(* Logix 5000 project; controller TFF vendor 1 type 14 code 107 rev 33.11; software revision 33.04; part 21 of 38 *)
(* tags used below, declared in another part *)
   Config : Configuration;   // Index Array used in configuration routines
   TIME : DINT[2];
   AA008 : ALIAS FOR DigitalPoint[18];
   AI101_SIG : ALIAS FOR DigitalPoint[106];
   AI104_SIG : ALIAS FOR DigitalPoint[107];
   AI201A_SIG : ALIAS FOR DigitalPoint[90];
   AI201B_SIG : ALIAS FOR DigitalPoint[109];
   AI202_SIG : ALIAS FOR DigitalPoint[105];
   AI203_SIG : ALIAS FOR DigitalPoint[91];
   AI204_SIG : ALIAS FOR DigitalPoint[92];
   DF24VDC : ALIAS FOR DigitalPoint[4];
   DF24VDCPC : ALIAS FOR DigitalPoint[25];
   DF3PHP003 : ALIAS FOR DigitalPoint[27];
   DF48MIX : ALIAS FOR DigitalPoint[26];
   DF48P001 : ALIAS FOR DigitalPoint[23];
   DF48P002 : ALIAS FOR DigitalPoint[24];
   Diafiltration : Diafiltration;
   DigitalPoint : DigitalPoint[150];   // Digital Point Array
   Drive : Drive[11];   // Drives Array
   ES001 : ALIAS FOR DigitalPoint[2];
   ExternalTCU : BOOL;   // Use of External TCU
   ExternalWeight : BOOL;   // Use of External Weight
   FI101_SIG : ALIAS FOR DigitalPoint[110];
   FI201_SIG : ALIAS FOR DigitalPoint[93];
   FI401_SIG : ALIAS FOR DigitalPoint[94];
   FlowPath : FlowPath[64];   // Flow Path Array
   FlowPathControl : FlowPathControl;   // Flow Path Control
   Gateway : Gateway;   // Gateway Control
   MIX101 : ALIAS FOR AnalogPoint[14];
   MIX101_SIG : ALIAS FOR DigitalPoint[104];
   MIX101DF : ALIAS FOR DigitalPoint[28];
   Mixer : Mixer;   // Mixer config. structure
   Options : Options;   // Options List
   PCV101 : ALIAS FOR AnalogPoint[3];
   PCV101_SIG : ALIAS FOR DigitalPoint[102];
   PCV201 : ALIAS FOR AnalogPoint[4];
   PCV201_SIG : ALIAS FOR DigitalPoint[103];
   PI001_SIG : ALIAS FOR DigitalPoint[97];
   PI101_SIG : ALIAS FOR DigitalPoint[98];
   PI201_SIG : ALIAS FOR DigitalPoint[99];
   PI401_SIG : ALIAS FOR DigitalPoint[100];
   PI601_SIG : ALIAS FOR DigitalPoint[95];
   PISL601 : ALIAS FOR DigitalPoint[0];
   PISL602 : ALIAS FOR DigitalPoint[1];
   PSH001 : ALIAS FOR DigitalPoint[21];
   PSH401 : ALIAS FOR DigitalPoint[22];
   RSBUZZ : ALIAS FOR DigitalPoint[3];
   SIC001 : ALIAS FOR Drive[1];
   SIC001DF : ALIAS FOR DigitalPoint[16];
   SIC002 : ALIAS FOR Drive[2];
   SIC002DF : ALIAS FOR DigitalPoint[17];
   SIC003DF : ALIAS FOR DigitalPoint[29];
   SIC004 : ALIAS FOR Drive[3];
   Tank : TankManagement;   // Tank Management
   TCU101_SIG : ALIAS FOR DigitalPoint[108];
   TCU101DF : ALIAS FOR DigitalPoint[30];
   TI101_SIG : ALIAS FOR DigitalPoint[101];
   TI201_SIG : ALIAS FOR DigitalPoint[111];
   UserCr1 : ALIAS FOR DigitalPoint[65];
   UserCr2 : ALIAS FOR DigitalPoint[67];
   UserNCr1 : ALIAS FOR DigitalPoint[64];
   UserNCr2 : ALIAS FOR DigitalPoint[66];
   Valve : Valve[100];   // Valve Array
   WI201_SIG : ALIAS FOR DigitalPoint[96];
   XS011 : ALIAS FOR DigitalPoint[14];
   XS012 : ALIAS FOR DigitalPoint[15];
   XV003 : ALIAS FOR Valve[2];
   YA01 : ALIAS FOR DigitalPoint[50];
   YA02 : ALIAS FOR DigitalPoint[51];
   YA03 : ALIAS FOR DigitalPoint[52];
   YA04 : ALIAS FOR DigitalPoint[53];
   YA05 : ALIAS FOR DigitalPoint[54];
   YA06 : ALIAS FOR DigitalPoint[55];
   YA07 : ALIAS FOR DigitalPoint[56];
   YA08 : ALIAS FOR DigitalPoint[57];
   YA09 : ALIAS FOR DigitalPoint[58];
   YA10 : ALIAS FOR DigitalPoint[59];
   YA11 : ALIAS FOR DigitalPoint[60];
   YA12 : ALIAS FOR DigitalPoint[61];
   YA13 : ALIAS FOR DigitalPoint[62];
   YA14 : ALIAS FOR DigitalPoint[63];
   YA15 : ALIAS FOR DigitalPoint[69];
   YA16 : ALIAS FOR DigitalPoint[70];
   YA17 : ALIAS FOR DigitalPoint[71];
   YA18 : ALIAS FOR DigitalPoint[72];
   YA41 : ALIAS FOR DigitalPoint[73];
   ZS001 : ALIAS FOR DigitalPoint[6];
   ZS002 : ALIAS FOR DigitalPoint[7];
   ZS003 : ALIAS FOR DigitalPoint[8];
   ZS004 : ALIAS FOR DigitalPoint[9];
   ZS005 : ALIAS FOR DigitalPoint[10];
   ZS008 : ALIAS FOR DigitalPoint[5];
   ZSDF : ALIAS FOR DigitalPoint[68];
(* Process, continued *)

ROUTINE Config_DigitalPoint_Real   (* structured text *)
// Apply the default configuration
   (* ==========================================================
   	Config DigitalPoint Real : Configure DigitalPoint Structure (for real input)
   
   	List of treatments
   		- DigitalPoint[0] : Valves Air Defect PISL601
   		- DigitalPoint[1] : Manifold Valves Air Defect PISL602
   		- DigitalPoint[2] : Emergency Stop ES001
   		- DigitalPoint[3] : Reset Buzzer RSBUZZ
   		- DigitalPoint[4] : 24 VDC defect DF24VDC
   		- DigitalPoint[5] : Door Closed ZS008
   		- DigitalPoint[6] : Clamshell Locking 1 Closed ZS001
   		- DigitalPoint[7] : Clamshell Locking 2 Closed ZS002
   		- DigitalPoint[8] : Clamshell Locking 3 Closed ZS003
   		- DigitalPoint[9] : Clamshell Locking 4 Closed ZS004
   		- DigitalPoint[10]: Clamshell Locking 5 Closed ZS005
   		- Reset Loop : Set to 0 the DigitalPoint[11 to 13].EnableCfg
   		- DigitalPoint[14]: Pump P001 Type XS011
   		- DigitalPoint[15]: Pump P002 Type XS012
   		- DigitalPoint[16]: P001 Defect SIC001DF
   		- DigitalPoint[17]: P002 Defect SIC002DF
   		- DigitalPoint[18]: C8000 Defect AA008
   		- DigitalPoint[19]: Spare
   		- DigitalPoint[20]: Spare
   		- DigitalPoint[21]: Feed Pump High Pressure PSH001
   		- DigitalPoint[22]: Transfer Pump High Pressure PSH401
   		- DigitalPoint[23]: P001 48 VDC Defect DF48P001
   		- DigitalPoint[24]: P002 48 VDC Defect DF48P002
   		- DigitalPoint[25]: Pump Cart 24 VDC Defect DF24VDCPC
   		- DigitalPoint[26]: Mixer 48 VDC Defect DF48MIX
   		- DigitalPoint[27]: Pump P003 Power Supply Defect DF3PHP003
   		- DigitalPoint[28]: Mixer Defect MIX101DF
   		- DigitalPoint[29]: P003 Defect SIC003DF
   		- DigitalPoint[30]: TCU Defect TCU101DF
   		- Reset Loop : Set to 0 the DigitalPoint[31 to 33].EnableCfg
   		- DigitalPoint[34]: Exchange DI#1
   		- DigitalPoint[35]: Exchange DI#2
   		- DigitalPoint[36]: Exchange DI#3
   		- DigitalPoint[37]: Exchange DI#4
   		- DigitalPoint[38]: Exchange DI#5
   		- DigitalPoint[39]: Exchange DI#6
   		- DigitalPoint[40]: Exchange DI#7
   		- DigitalPoint[41]: Exchange DI#8
   		- Reset Loop : Set to 0 the DigitalPoint[42 to 49].EnableCfg
   
   -----------------------------------------------------------------------------------------------------------------------------------------------------
   	History
   		2019-DEC-24 - Merck - Q. Spindler - Initial version for Candidate Release 1.00.00.00.a
   		2020-MAR-27 - Merck - Q. Spindler - Modifications for Candidate Release 1.00.00.00.b
   					- Add Options for AA008
   		2020-SEP-09 - Merck - Q. Spindler - Modifications for Candidate Release 1.00.00.00.d
   					- Change PriorityCfg to 0 and set Priority to 1 for PSH001 and PSH401
   					- Disable TCU101DF alarm if ExternalTCU not used
   ============================================================*)
   
   (*DigitalPoint[0] : Valves Air Defect PISL601
   ============================================================*)
   DigitalPoint[0].EnableCfg := 1 ;
   DigitalPoint[0].ActiveStateCFg := 1 ;
   DigitalPoint[0].RealInputCfg := 1 ;
   DigitalPoint[0].InputAddressCfg := 0 ;
   DigitalPoint[0].AlarmCfg := 1 ;
   DigitalPoint[0].AlarmStateCfg := 0 ;
   DigitalPoint[0].OverrideCfg := 1 ;
   DigitalPoint[0].PriorityCfg := 1 ;
   DigitalPoint[0].Cond1Cfg := 0 ;
   DigitalPoint[0].Cond2Cfg := 0 ;
   DigitalPoint[0].FlashingInputCfg := 0 ;
   
   (*DigitalPoint[1] : Manifold Valves Air Defect PISL602
   ============================================================*)
   DigitalPoint[1].EnableCfg := 1 ;
   DigitalPoint[1].ActiveStateCFg := 1 ;
   DigitalPoint[1].RealInputCfg := 1 ;
   DigitalPoint[1].InputAddressCfg := 1 ;
   DigitalPoint[1].AlarmCfg := 1 ;
   DigitalPoint[1].AlarmStateCfg := 0 ;
   DigitalPoint[1].OverrideCfg := 1 ;
   DigitalPoint[1].PriorityCfg := 1 ;
   DigitalPoint[1].Cond1Cfg := 0 ;
   DigitalPoint[1].Cond2Cfg := 0 ;
   DigitalPoint[1].FlashingInputCfg := 0 ;
   
   (*DigitalPoint[2] : Emergency Stop ES001
   ============================================================*)
   DigitalPoint[2].EnableCfg := 1 ;
   DigitalPoint[2].ActiveStateCFg := 1 ;
   DigitalPoint[2].RealInputCfg := 1 ;
   DigitalPoint[2].InputAddressCfg := 2 ;
   DigitalPoint[2].AlarmCfg := 1 ;
   DigitalPoint[2].AlarmStateCfg := 0 ;
   DigitalPoint[2].OverrideCfg := 0 ;
   DigitalPoint[2].PriorityCfg := 0 ;
   DigitalPoint[2].Priority := 1 ;
   DigitalPoint[2].Cond1Cfg := 0 ;
   DigitalPoint[2].Cond2Cfg := 0 ;
   DigitalPoint[2].FlashingInputCfg := 0 ;
   
   (*DigitalPoint[3] : Reset Buzzer RSBUZZ
   ============================================================*)
   DigitalPoint[3].EnableCfg := 1 ;
   DigitalPoint[3].ActiveStateCFg := 1 ;
   DigitalPoint[3].RealInputCfg := 1 ;
   DigitalPoint[3].InputAddressCfg := 3 ;
   DigitalPoint[3].AlarmCfg := 0 ;
   DigitalPoint[3].Alarm := 0 ;
   DigitalPoint[3].AlarmStateCfg := 0 ;
   DigitalPoint[3].OverrideCfg := 0 ;
   DigitalPoint[3].Priority := 0 ;
   DigitalPoint[3].PriorityCfg := 0 ;
   DigitalPoint[3].Cond1Cfg := 0 ;
   DigitalPoint[3].Cond2Cfg := 0 ;
   DigitalPoint[3].FlashingInputCfg := 0 ;
   
   (*DigitalPoint[4] : 24 VDC defect DF24VDC
   ============================================================*)
   DigitalPoint[4].EnableCfg := 1 ;
   DigitalPoint[4].ActiveStateCFg := 1 ;
   DigitalPoint[4].RealInputCfg := 1 ;
   DigitalPoint[4].InputAddressCfg := 4 ;
   DigitalPoint[4].AlarmCfg := 1 ;
   DigitalPoint[4].AlarmStateCfg := 0 ;
   DigitalPoint[4].OverrideCfg := 1 ;
   DigitalPoint[4].PriorityCfg := 1 ;
   DigitalPoint[4].Cond1Cfg := 0 ;
   DigitalPoint[4].Cond2Cfg := 0 ;
   DigitalPoint[4].FlashingInputCfg := 0 ;
   
   (*DigitalPoint[5] : Door Closed ZS008
   ============================================================*)
   DigitalPoint[5].EnableCfg := 1 ;
   DigitalPoint[5].ActiveStateCFg := 1 ;
   DigitalPoint[5].RealInputCfg := 1 ;
   DigitalPoint[5].InputAddressCfg := 5 ;
   DigitalPoint[5].AlarmCfg := 1 ;
   DigitalPoint[5].AlarmStateCfg := 0 ;
   DigitalPoint[5].OverrideCfg := 1 ;
   DigitalPoint[5].PriorityCfg := 1 ;
   DigitalPoint[5].Cond1Cfg := 0 ;
   DigitalPoint[5].Cond2Cfg := 0 ;
   DigitalPoint[5].FlashingInputCfg := 0 ;
   
   (*DigitalPoint[6] : Clamshell Locking 1 Closed ZS001
   ============================================================*)
   DigitalPoint[6].EnableCfg := 1 ;
   DigitalPoint[6].ActiveStateCFg := 1 ;
   DigitalPoint[6].RealInputCfg := 1 ;
   DigitalPoint[6].InputAddressCfg := 6 ;
   DigitalPoint[6].AlarmCfg := 0 ;
   DigitalPoint[6].Alarm := 0 ;
   DigitalPoint[6].AlarmStateCfg := 0 ;
   DigitalPoint[6].OverrideCfg := 0 ;
   DigitalPoint[6].PriorityCfg := 0 ;
   DigitalPoint[6].Cond1Cfg := 0 ;
   DigitalPoint[6].Cond2Cfg := 0 ;
   DigitalPoint[6].FlashingInputCfg := 0 ;
   
   (*DigitalPoint[7] : Clamshell Locking 2 Closed ZS002
   ============================================================*)
   DigitalPoint[7].EnableCfg := 1 ;
   DigitalPoint[7].ActiveStateCFg := 1 ;
   DigitalPoint[7].RealInputCfg := 1 ;
   DigitalPoint[7].InputAddressCfg := 7 ;
   DigitalPoint[7].AlarmCfg := 0 ;
   DigitalPoint[7].Alarm := 0 ;
   DigitalPoint[7].AlarmStateCfg := 0 ;
   DigitalPoint[7].OverrideCfg := 0 ;
   DigitalPoint[7].PriorityCfg := 0 ;
   DigitalPoint[7].Cond1Cfg := 0 ;
   DigitalPoint[7].Cond2Cfg := 0 ;
   DigitalPoint[7].FlashingInputCfg := 0 ;
   
   (*DigitalPoint[8] : Clamshell Locking 3 Closed ZS003
   ============================================================*)
   DigitalPoint[8].EnableCfg := 1 ;
   DigitalPoint[8].ActiveStateCFg := 1 ;
   DigitalPoint[8].RealInputCfg := 1 ;
   DigitalPoint[8].InputAddressCfg := 8 ;
   DigitalPoint[8].AlarmCfg := 0 ;
   DigitalPoint[8].Alarm := 0 ;
   DigitalPoint[8].AlarmStateCfg := 0 ;
   DigitalPoint[8].OverrideCfg := 0 ;
   DigitalPoint[8].PriorityCfg := 0 ;
   DigitalPoint[8].Cond1Cfg := 0 ;
   DigitalPoint[8].Cond2Cfg := 0 ;
   DigitalPoint[8].FlashingInputCfg := 0 ;
   
   (*DigitalPoint[9] : Clamshell Locking 4 Closed ZS004
   ============================================================*)
   DigitalPoint[9].EnableCfg := 1 ;
   DigitalPoint[9].ActiveStateCFg := 1 ;
   DigitalPoint[9].RealInputCfg := 1 ;
   DigitalPoint[9].InputAddressCfg := 9 ;
   DigitalPoint[9].AlarmCfg := 0 ;
   DigitalPoint[9].Alarm := 0 ;
   DigitalPoint[9].AlarmStateCfg := 0 ;
   DigitalPoint[9].OverrideCfg := 0 ;
   DigitalPoint[9].PriorityCfg := 0 ;
   DigitalPoint[9].Cond1Cfg := 0 ;
   DigitalPoint[9].Cond2Cfg := 0 ;
   DigitalPoint[9].FlashingInputCfg := 0 ;
   
   (*DigitalPoint[10]: Clamshell Locking 5 Closed ZS005
   ============================================================*)
   DigitalPoint[10].EnableCfg := 1 ;
   DigitalPoint[10].ActiveStateCFg := 1 ;
   DigitalPoint[10].RealInputCfg := 1 ;
   DigitalPoint[10].InputAddressCfg := 10 ;
   DigitalPoint[10].AlarmCfg := 0 ;
   DigitalPoint[10].Alarm := 0 ;
   DigitalPoint[10].AlarmStateCfg := 0 ;
   DigitalPoint[10].OverrideCfg := 0 ;
   DigitalPoint[10].PriorityCfg := 0 ;
   DigitalPoint[10].Cond1Cfg := 0 ;
   DigitalPoint[10].Cond2Cfg := 0 ;
   DigitalPoint[10].FlashingInputCfg := 0 ;
   
   
   (*Reset Loop : Set to 0 the DigitalPoint[11 to 13].EnableCfg
   ============================================================*)
   FOR Config.IndexDP := 11 to 13 do
   	DigitalPoint[Config.IndexDP].EnableCfg := 0 ;
   	DigitalPoint[Config.IndexDP].AlarmCfg := 0 ;
   	DigitalPoint[Config.IndexDP].Alarm := 0 ;
   End_for ;
   
   
   (*DigitalPoint[14]: Pump P001 Type XS011
   ============================================================*)
   DigitalPoint[14].EnableCfg := 1 ;
   DigitalPoint[14].ActiveStateCFg := 1 ;
   DigitalPoint[14].RealInputCfg := 1 ;
   DigitalPoint[14].InputAddressCfg := 14 ;
   DigitalPoint[14].AlarmCfg := 0 ;
   DigitalPoint[14].Alarm := 0 ;
   DigitalPoint[14].AlarmStateCfg := 0 ;
   DigitalPoint[14].OverrideCfg := 0 ;
   DigitalPoint[14].PriorityCfg := 0 ;
   DigitalPoint[14].Cond1Cfg := 0 ;
   DigitalPoint[14].Cond2Cfg := 0 ;
   DigitalPoint[14].FlashingInputCfg := 0 ;
   
   (*DigitalPoint[15]: Pump P002 Type XS012
   ============================================================*)
   DigitalPoint[15].EnableCfg := 1 ;
   DigitalPoint[15].ActiveStateCFg := 1 ;
   DigitalPoint[15].RealInputCfg := 1 ;
   DigitalPoint[15].InputAddressCfg := 15 ;
   DigitalPoint[15].AlarmCfg := 0 ;
   DigitalPoint[15].Alarm := 0 ;
   DigitalPoint[15].AlarmStateCfg := 0 ;
   DigitalPoint[15].OverrideCfg := 0 ;
   DigitalPoint[15].PriorityCfg := 0 ;
   DigitalPoint[15].Cond1Cfg := 0 ;
   DigitalPoint[15].Cond2Cfg := 0 ;
   DigitalPoint[15].FlashingInputCfg := 0 ;
   
   (*DigitalPoint[16]: P001 Defect SIC001DF
   ============================================================*)
   DigitalPoint[16].EnableCfg := 1 ;
   DigitalPoint[16].ActiveStateCFg := 1 ;
   DigitalPoint[16].RealInputCfg := 1 ;
   DigitalPoint[16].InputAddressCfg := 16 ;
   DigitalPoint[16].AlarmCfg := 1 ;
   DigitalPoint[16].AlarmStateCfg := 0 ;
   DigitalPoint[16].OverrideCfg := 1 ;
   DigitalPoint[16].PriorityCfg := 1 ;
   DigitalPoint[16].Cond1Cfg := 0 ;
   DigitalPoint[16].Cond2Cfg := 0 ;
   DigitalPoint[16].FlashingInputCfg := 0 ;
   
   (*DigitalPoint[17]: P002 Defect SIC002DF
   ============================================================*)
   DigitalPoint[17].EnableCfg := 1 ;
   DigitalPoint[17].ActiveStateCFg := 1 ;
   DigitalPoint[17].RealInputCfg := 1 ;
   DigitalPoint[17].InputAddressCfg := 17 ;
   DigitalPoint[17].AlarmCfg := 1 ;
   DigitalPoint[17].AlarmStateCfg := 0 ;
   DigitalPoint[17].OverrideCfg := 1 ;
   DigitalPoint[17].PriorityCfg := 1 ;
   DigitalPoint[17].Cond1Cfg := 0 ;
   DigitalPoint[17].Cond2Cfg := 0 ;
   DigitalPoint[17].FlashingInputCfg := 0 ;
   
   (*DigitalPoint[18]: C8000 Defect AA008
   ============================================================*)
   If Options.FiltrateCondPHUV OR Options.FiltrateCondPH Then
   	DigitalPoint[18].EnableCfg := 1 ;
   	DigitalPoint[18].AlarmCfg := 1 ;
   Else
   	DigitalPoint[18].EnableCfg := 0 ;
   	DigitalPoint[18].AlarmCfg := 0 ;
   	DigitalPoint[18].Alarm := 0 ;
   End_if;
   
   DigitalPoint[18].ActiveStateCFg := 1 ;
   DigitalPoint[18].RealInputCfg := 1 ;
   DigitalPoint[18].InputAddressCfg := 18 ;
   DigitalPoint[18].AlarmStateCfg := 0 ;
   DigitalPoint[18].OverrideCfg := 1 ;
   DigitalPoint[18].PriorityCfg := 1 ;
   DigitalPoint[18].Cond1Cfg := 0 ;
   DigitalPoint[18].Cond2Cfg := 0 ;
   DigitalPoint[18].FlashingInputCfg := 0 ;
   
   (*DigitalPoint[19]: Spare
   ============================================================*)
   DigitalPoint[19].EnableCfg := 0 ;
   DigitalPoint[19].ActiveStateCFg := 1 ;
   DigitalPoint[19].RealInputCfg := 1 ;
   DigitalPoint[19].InputAddressCfg := 19 ;
   DigitalPoint[19].AlarmCfg := 0 ;
   DigitalPoint[19].AlarmStateCfg := 0 ;
   DigitalPoint[19].OverrideCfg := 1 ;
   DigitalPoint[19].PriorityCfg := 1 ;
   DigitalPoint[19].Cond1Cfg := 0 ;
   DigitalPoint[19].Cond2Cfg := 0 ;
   DigitalPoint[19].FlashingInputCfg := 0 ;
   
   (*DigitalPoint[20]: Spare
   ============================================================*)
   DigitalPoint[20].EnableCfg := 0 ;
   DigitalPoint[20].ActiveStateCFg := 1 ;
   DigitalPoint[20].RealInputCfg := 1 ;
   DigitalPoint[20].InputAddressCfg := 20 ;
   DigitalPoint[20].AlarmCfg := 0 ;
   DigitalPoint[20].AlarmStateCfg := 0 ;
   DigitalPoint[20].OverrideCfg := 1 ;
   DigitalPoint[20].PriorityCfg := 1 ;
   DigitalPoint[20].Cond1Cfg := 0 ;
   DigitalPoint[20].Cond2Cfg := 0 ;
   DigitalPoint[20].FlashingInputCfg := 0 ;
   
   (*DigitalPoint[21]: Feed Pump High Pressure PSH001
   ============================================================*)
   DigitalPoint[21].EnableCfg := 1 ;
   DigitalPoint[21].ActiveStateCFg := 1 ;
   DigitalPoint[21].RealInputCfg := 1 ;
   DigitalPoint[21].InputAddressCfg := 21 ;
   DigitalPoint[21].AlarmCfg := 1 ;
   DigitalPoint[21].AlarmStateCfg := 0 ;
   DigitalPoint[21].OverrideCfg := 1 ;
   DigitalPoint[21].PriorityCfg := 0 ;
   DigitalPoint[21].Priority := 1 ;
   DigitalPoint[21].Cond1Cfg := 0 ;
   DigitalPoint[21].Cond2Cfg := 0 ;
   DigitalPoint[21].FlashingInputCfg := 0 ;
   
   (*DigitalPoint[22]: Transfer Pump High Pressure PSH401
   ============================================================*)
   DigitalPoint[22].EnableCfg := 1 ;
   DigitalPoint[22].ActiveStateCFg := 1 ;
   DigitalPoint[22].RealInputCfg := 1 ;
   DigitalPoint[22].InputAddressCfg := 22 ;
   DigitalPoint[22].AlarmCfg := 1 ;
   DigitalPoint[22].AlarmStateCfg := 0 ;
   DigitalPoint[22].OverrideCfg := 1 ;
   DigitalPoint[22].PriorityCfg := 0 ;
   DigitalPoint[22].Priority := 1 ;
   DigitalPoint[22].Cond1Cfg := 0 ;
   DigitalPoint[22].Cond2Cfg := 0 ;
   DigitalPoint[22].FlashingInputCfg := 0 ;
   
   (*DigitalPoint[23]: P001 48 VDC Defect DF48P001
   ============================================================*)
   DigitalPoint[23].EnableCfg := 1 ;
   DigitalPoint[23].ActiveStateCFg := 1 ;
   DigitalPoint[23].RealInputCfg := 1 ;
   DigitalPoint[23].InputAddressCfg := 23 ;
   DigitalPoint[23].AlarmCfg := 1 ;
   DigitalPoint[23].AlarmStateCfg := 0 ;
   DigitalPoint[23].OverrideCfg := 1 ;
   DigitalPoint[23].PriorityCfg := 1 ;
   DigitalPoint[23].Cond1Cfg := 0 ;
   DigitalPoint[23].Cond2Cfg := 0 ;
   DigitalPoint[23].FlashingInputCfg := 0 ;
   
   (*DigitalPoint[24]: P002 48 VDC Defect DF48P002
   ============================================================*)
   DigitalPoint[24].EnableCfg := 1 ;
   DigitalPoint[24].ActiveStateCFg := 1 ;
   DigitalPoint[24].RealInputCfg := 1 ;
   DigitalPoint[24].InputAddressCfg := 24 ;
   DigitalPoint[24].AlarmCfg := 1 ;
   DigitalPoint[24].AlarmStateCfg := 0 ;
   DigitalPoint[24].OverrideCfg := 1 ;
   DigitalPoint[24].PriorityCfg := 1 ;
   DigitalPoint[24].Cond1Cfg := 0 ;
   DigitalPoint[24].Cond2Cfg := 0 ;
   DigitalPoint[24].FlashingInputCfg := 0 ;
   
   (*DigitalPoint[25]: Pump Cart 24 VDC Defect DF24VDCPC
   ============================================================*)
   DigitalPoint[25].EnableCfg := 1 ;
   DigitalPoint[25].ActiveStateCFg := 1 ;
   DigitalPoint[25].RealInputCfg := 1 ;
   DigitalPoint[25].InputAddressCfg := 25 ;
   DigitalPoint[25].AlarmCfg := 1 ;
   DigitalPoint[25].AlarmStateCfg := 0 ;
   DigitalPoint[25].OverrideCfg := 1 ;
   DigitalPoint[25].PriorityCfg := 1 ;
   DigitalPoint[25].Cond1Cfg := 0 ;
   DigitalPoint[25].Cond2Cfg := 0 ;
   DigitalPoint[25].FlashingInputCfg := 0 ;
   
   (*DigitalPoint[26]: Mixer 48 VDC Defect DF48MIX
   ============================================================*)
   (*Set to 1 to use this DigitalPoint*)
   If Options.FeedTank then
   	DigitalPoint[26].EnableCfg := 1 ;
   	DigitalPoint[26].AlarmCfg := 1 ;
   else
   	DigitalPoint[26].EnableCfg := 0 ;
   	DigitalPoint[26].AlarmCfg := 0 ;
   	DigitalPoint[26].Alarm := 0 ;
   End_if;
   DigitalPoint[26].ActiveStateCFg := 1 ;
   DigitalPoint[26].RealInputCfg := 1 ;
   DigitalPoint[26].InputAddressCfg := 26 ;
   DigitalPoint[26].AlarmStateCfg := 0 ;
   DigitalPoint[26].OverrideCfg := 1 ;
   DigitalPoint[26].PriorityCfg := 1 ;
   DigitalPoint[26].Cond1Cfg := 0 ;
   DigitalPoint[26].Cond2Cfg := 0 ;
   DigitalPoint[26].FlashingInputCfg := 0 ;
   
   (*DigitalPoint[27]: Pump P003 Power Supply Defect DF3PHP003
   ============================================================*)
   DigitalPoint[27].EnableCfg := 1 ;
   DigitalPoint[27].ActiveStateCFg := 1 ;
   DigitalPoint[27].RealInputCfg := 1 ;
   DigitalPoint[27].InputAddressCfg := 27 ;
   DigitalPoint[27].AlarmCfg := 1 ;
   DigitalPoint[27].AlarmStateCfg := 0 ;
   DigitalPoint[27].OverrideCfg := 1 ;
   DigitalPoint[27].PriorityCfg := 1 ;
   DigitalPoint[27].Cond1Cfg := 0 ;
   DigitalPoint[27].Cond2Cfg := 0 ;
   DigitalPoint[27].FlashingInputCfg := 0 ;
   
   (*DigitalPoint[28]: Mixer Defect MIX101DF
   ============================================================*)
   (*Set to 1 to use this DigitalPoint*)
   If Options.FeedTank then
   	DigitalPoint[28].EnableCfg := 1 ;
   	DigitalPoint[28].AlarmCfg := 1 ;
   else
   	DigitalPoint[28].EnableCfg := 0 ;
   	DigitalPoint[28].AlarmCfg := 0 ;
   	DigitalPoint[28].Alarm := 0 ;
   End_if;
   DigitalPoint[28].ActiveStateCFg := 1 ;
   DigitalPoint[28].RealInputCfg := 1 ;
   DigitalPoint[28].InputAddressCfg := 28 ;
   DigitalPoint[28].AlarmStateCfg := 0 ;
   DigitalPoint[28].OverrideCfg := 1 ;
   DigitalPoint[28].PriorityCfg := 1 ;
   DigitalPoint[28].Cond1Cfg := 0 ;
   DigitalPoint[28].Cond2Cfg := 0 ;
   DigitalPoint[28].FlashingInputCfg := 0 ;
   
   (*DigitalPoint[29]: P003 Defect SIC003DF
   ============================================================*)
   DigitalPoint[29].EnableCfg := 1 ;
   DigitalPoint[29].ActiveStateCFg := 1 ;
   DigitalPoint[29].RealInputCfg := 1 ;
   DigitalPoint[29].InputAddressCfg := 29 ;
   DigitalPoint[29].AlarmCfg := 1 ;
   DigitalPoint[29].AlarmStateCfg := 0 ;
   DigitalPoint[29].OverrideCfg := 1 ;
   DigitalPoint[29].PriorityCfg := 1 ;
   DigitalPoint[29].Cond1Cfg := 0 ;
   DigitalPoint[29].Cond2Cfg := 0 ;
   DigitalPoint[29].FlashingInputCfg := 0 ;
   
   (*DigitalPoint[30]: TCU Defect TCU101DF
   ============================================================*)
   (*Set to 1 to use this DigitalPoint*)
   If Options.FeedTank then
   	DigitalPoint[30].EnableCfg := 1 ;
   	If ExternalTCU then
   		DigitalPoint[30].AlarmCfg := 1 ;
   	else
   		DigitalPoint[30].AlarmCfg := 0 ;
   		DigitalPoint[30].Alarm := 0 ;
   	End_if;
   else
   	DigitalPoint[30].EnableCfg := 0 ;
   	DigitalPoint[30].AlarmCfg := 0 ;
   	DigitalPoint[30].Alarm := 0 ;
   End_if;
   DigitalPoint[30].ActiveStateCFg := 1 ;
   DigitalPoint[30].RealInputCfg := 1 ;
   DigitalPoint[30].InputAddressCfg := 30 ;
   DigitalPoint[30].AlarmStateCfg := 0 ;
   DigitalPoint[30].OverrideCfg := 1 ;
   DigitalPoint[30].PriorityCfg := 1 ;
   DigitalPoint[30].Cond1Cfg := 0 ;
   DigitalPoint[30].Cond2Cfg := 0 ;
   DigitalPoint[30].FlashingInputCfg := 0 ;
   
   (*Reset Loop : Set to 0 the DigitalPoint[31 to 33].EnableCfg
   ============================================================*)
   FOR Config.IndexDP := 31 to 33 do
   	DigitalPoint[Config.IndexDP].EnableCfg := 0 ;
   	DigitalPoint[Config.IndexDP].AlarmCfg := 0 ;
   	DigitalPoint[Config.IndexDP].Alarm := 0 ;
   End_for ;
   
   (*DigitalPoint[34]: Exchange DI#1
   ============================================================*)
   (*Set to 1 to use this DigitalPoint*)
   If Options.External_IO then
   	DigitalPoint[34].EnableCfg := 1 ;
   else
   	DigitalPoint[34].EnableCfg := 0 ;
   End_if ;
   (*Default Configuration *)
   DigitalPoint[34].ActiveStateCFg := 1 ;
   DigitalPoint[34].RealInputCfg := 1 ;
   DigitalPoint[34].InputAddressCfg := 34 ;
   DigitalPoint[34].AlarmStateCfg := 0 ;
   DigitalPoint[34].OverrideCfg := 0 ;
   DigitalPoint[34].PriorityCfg := 0 ;
   DigitalPoint[34].Cond1Cfg := 0 ;
   DigitalPoint[34].Cond2Cfg := 0 ;
   DigitalPoint[34].FlashingInputCfg := 0 ;
   DigitalPoint[34].AlarmCfg := 0 ;
   
   (*DigitalPoint[35]: Exchange DI#2
   ============================================================*)
   (*Set to 1 to use this DigitalPoint*)
   If Options.External_IO then
   	DigitalPoint[35].EnableCfg := 1 ;
   else
   	DigitalPoint[35].EnableCfg := 0 ;
   End_if ;
   (*Default Configuration *)
   DigitalPoint[35].ActiveStateCFg := 1 ;
   DigitalPoint[35].RealInputCfg := 1 ;
   DigitalPoint[35].InputAddressCfg := 35 ;
   DigitalPoint[35].AlarmStateCfg := 0 ;
   DigitalPoint[35].OverrideCfg := 0 ;
   DigitalPoint[35].PriorityCfg := 0 ;
   DigitalPoint[35].Cond1Cfg := 0 ;
   DigitalPoint[35].Cond2Cfg := 0 ;
   DigitalPoint[35].FlashingInputCfg := 0 ;
   DigitalPoint[35].AlarmCfg := 0 ;
   
   (*DigitalPoint[36]: Exchange DI#3
   ============================================================*)
   (*Set to 1 to use this DigitalPoint*)
   If Options.External_IO then
   	DigitalPoint[36].EnableCfg := 1 ;
   else
   	DigitalPoint[36].EnableCfg := 0 ;
   End_if ;
   (*Default Configuration *)
   DigitalPoint[36].ActiveStateCFg := 1 ;
   DigitalPoint[36].RealInputCfg := 1 ;
   DigitalPoint[36].InputAddressCfg := 36 ;
   DigitalPoint[36].AlarmStateCfg := 0 ;
   DigitalPoint[36].OverrideCfg := 0 ;
   DigitalPoint[36].PriorityCfg := 0 ;
   DigitalPoint[36].Cond1Cfg := 0 ;
   DigitalPoint[36].Cond2Cfg := 0 ;
   DigitalPoint[36].FlashingInputCfg := 0 ;
   DigitalPoint[36].AlarmCfg := 0 ;
   
   (*DigitalPoint[37]: Exchange DI#4
   ============================================================*)
   (*Set to 1 to use this DigitalPoint*)
   If Options.External_IO then
   	DigitalPoint[37].EnableCfg := 1 ;
   else
   	DigitalPoint[37].EnableCfg := 0 ;
   End_if ;
   (*Default Configuration *)
   DigitalPoint[37].ActiveStateCFg := 1 ;
   DigitalPoint[37].RealInputCfg := 1 ;
   DigitalPoint[37].InputAddressCfg := 37 ;
   DigitalPoint[37].AlarmStateCfg := 0 ;
   DigitalPoint[37].OverrideCfg := 0 ;
   DigitalPoint[37].PriorityCfg := 0 ;
   DigitalPoint[37].Cond1Cfg := 0 ;
   DigitalPoint[37].Cond2Cfg := 0 ;
   DigitalPoint[37].FlashingInputCfg := 0 ;
   DigitalPoint[37].AlarmCfg := 0 ;
   
   (*DigitalPoint[38]: Exchange DI#5
   ============================================================*)
   (*Set to 1 to use this DigitalPoint*)
   If Options.External_IO then
   	DigitalPoint[38].EnableCfg := 1 ;
   else
   	DigitalPoint[38].EnableCfg := 0 ;
   End_if ;
   (*Default Configuration *)
   DigitalPoint[38].ActiveStateCFg := 1 ;
   DigitalPoint[38].RealInputCfg := 1 ;
   DigitalPoint[38].InputAddressCfg := 38 ;
   DigitalPoint[38].AlarmStateCfg := 0 ;
   DigitalPoint[38].OverrideCfg := 0 ;
   DigitalPoint[38].PriorityCfg := 0 ;
   DigitalPoint[38].Cond1Cfg := 0 ;
   DigitalPoint[38].Cond2Cfg := 0 ;
   DigitalPoint[38].FlashingInputCfg := 0 ;
   DigitalPoint[38].AlarmCfg := 0 ;
   
   (*DigitalPoint[39]: Exchange DI#6
   ============================================================*)
   (*Set to 1 to use this DigitalPoint*)
   If Options.External_IO then
   	DigitalPoint[39].EnableCfg := 1 ;
   else
   	DigitalPoint[39].EnableCfg := 0 ;
   End_if ;
   (*Default Configuration *)
   DigitalPoint[39].ActiveStateCFg := 1 ;
   DigitalPoint[39].RealInputCfg := 1 ;
   DigitalPoint[39].InputAddressCfg := 39 ;
   DigitalPoint[39].AlarmStateCfg := 0 ;
   DigitalPoint[39].OverrideCfg := 0 ;
   DigitalPoint[39].PriorityCfg := 0 ;
   DigitalPoint[39].Cond1Cfg := 0 ;
   DigitalPoint[39].Cond2Cfg := 0 ;
   DigitalPoint[39].FlashingInputCfg := 0 ;
   DigitalPoint[39].AlarmCfg := 0 ;
   
   (*DigitalPoint[40]: Exchange DI#7
   ============================================================*)
   (*Set to 1 to use this DigitalPoint*)
   If Options.External_IO then
   	DigitalPoint[40].EnableCfg := 1 ;
   else
   	DigitalPoint[40].EnableCfg := 0 ;
   End_if ;
   (*Default Configuration *)
   DigitalPoint[40].ActiveStateCFg := 1 ;
   DigitalPoint[40].RealInputCfg := 1 ;
   DigitalPoint[40].InputAddressCfg := 40 ;
   DigitalPoint[40].AlarmStateCfg := 0 ;
   DigitalPoint[40].OverrideCfg := 0 ;
   DigitalPoint[40].PriorityCfg := 0 ;
   DigitalPoint[40].Cond1Cfg := 0 ;
   DigitalPoint[40].Cond2Cfg := 0 ;
   DigitalPoint[40].FlashingInputCfg := 0 ;
   DigitalPoint[40].AlarmCfg := 0 ;
   
   (*DigitalPoint[41]: Exchange DI#8
   ============================================================*)
   (*Set to 1 to use this DigitalPoint*)
   If Options.External_IO then
   	DigitalPoint[41].EnableCfg := 1 ;
   else
   	DigitalPoint[41].EnableCfg := 0 ;
   End_if ;
   (*Default Configuration *)
   DigitalPoint[41].ActiveStateCFg := 1 ;
   DigitalPoint[41].RealInputCfg := 1 ;
   DigitalPoint[41].InputAddressCfg := 41 ;
   DigitalPoint[41].AlarmStateCfg := 0 ;
   DigitalPoint[41].OverrideCfg := 0 ;
   DigitalPoint[41].PriorityCfg := 0 ;
   DigitalPoint[41].Cond1Cfg := 0 ;
   DigitalPoint[41].Cond2Cfg := 0 ;
   DigitalPoint[41].FlashingInputCfg := 0 ;
   DigitalPoint[41].AlarmCfg := 0 ;
   
   (*Reset Loop : Set to 0 the DigitalPoint[42 to 49].EnableCfg
   ============================================================*)
   FOR Config.IndexDP := 42 to 49 do
   	DigitalPoint[Config.IndexDP].EnableCfg := 0 ;
   	DigitalPoint[Config.IndexDP].AlarmCfg := 0 ;
   	DigitalPoint[Config.IndexDP].Alarm := 0 ;
   End_for ;
END_ROUTINE

ROUTINE Config_DigitalPoint_Soft   (* structured text *)
   (* ==========================================================
   	Config DigitalPoint Soft : Configure DigitalPoint Structure (for soft input)
   
   	List of treatments
   		- DigitalPoint[50]: YA01 PC to PLC Com. Failure
   		- DigitalPoint[51]: YA02 CCP Runtime Com. Failure
   		- DigitalPoint[52]: YA03 Historical Data Collection Failure
   		- DigitalPoint[53]: YA04 Hard drive Overload
   		- DigitalPoint[54]: YA05 Database Overload
   		- DigitalPoint[55]: YA06 Node 0 Communication Failure - Smart
   		- DigitalPoint[56]: YA07 Node 0 Internal Defect - Smart
   		- DigitalPoint[57]: YA08 Node 1 Communication Failure - Clamshell
   		- DigitalPoint[58]: YA09 Node 1 Internal Defect - Clamshell
   		- DigitalPoint[59]: YA10 PLC Program Major Fault
   		- DigitalPoint[60]: YA11 Database Corrupted
   		- DigitalPoint[61]: YA12 Unauthorized accesses
   		- DigitalPoint[62]: YA13 Tank Size Mismatch
   		- DigitalPoint[63]: YA14 SQL Server Write Failure
   		- DigitalPoint[64]: UserNCr1 User Non Critical Alarm 1
   		- DigitalPoint[65]: UserCr1 User Critical Alarm 1
   		- DigitalPoint[66]: UserNCr2 User Non Critical Alarm 2
   		- DigitalPoint[67]: UserCr2 User Critical Alarm 2
   		- DigitalPoint[68]: ZSDF Clamshell Locking Defect
   		- DigitalPoint[69]: YA15 ACT350 Communication Failure
   		- DigitalPoint[70]: YA16 Watchdog Gateway
   		- DigitalPoint[71]: YA17 Mobius Device Communication Failure
   		- DigitalPoint[72]: YA18 Pump Type Mismatch
   		- DigitalPoint[73]: YA41 Operating Time Exceeded
   		- Reset Loop : Set to 0 the DigitalPoint[74 to 89].EnableCfg
   		- DigitalPoint[90]: AI201A_SIG Filtrate Conductivity Process Signal default
   		- DigitalPoint[91]: AI203_SIG Filtrate UV1 Signal default
   		- DigitalPoint[92]: AI204_SIG Filtrate UV2 Signal default
   		- DigitalPoint[93]: FI201_SIG Filtrate Flow Signal default
   		- DigitalPoint[94]: FI401_SIG Transfer Pump Flow Signal default
   		- DigitalPoint[95]: PI601_SIG Feed Tank Pressure Signal default
   		- DigitalPoint[96]: WI201_SIG External Filtrate Weight Signal default
   		- DigitalPoint[97]: PI001_SIG Feed Pressure Signal default
   		- DigitalPoint[98]: PI101_SIG Retentate Pressure Signal default
   		- DigitalPoint[99]: PI201_SIG Filtrate Pressure Signal default
   		- DigitalPoint[100]: PI401_SIG Transfer Pump Pressure Signal default
   		- DigitalPoint[101]: TI101_SIG Feed Tank Temperature Signal default
   		- DigitalPoint[102]: PCV101_SIG PCV101 Position Signal default
   		- DigitalPoint[103]: PCV201_SIG PCV201 Position Signal default
   		- DigitalPoint[104]: MIX101_SIG Mixer Speed Signal default
   		- DigitalPoint[105]: AI202_SIG Filtrate pH Signal default
   		- DigitalPoint[106]: AI101_SIG Feed Tank pH Signal default
   		- DigitalPoint[107]: AI104_SIG Feed Tank Conductivity Signal default
   		- DigitalPoint[108]: TCU101_SIG TCU Temperature Signal default
   		- DigitalPoint[109]: AI201B_SIG Filtrate Conductivity Cleaning Signal default
   		- DigitalPoint[110]: FI101_SIG Retentate Flow Signal default
   		- DigitalPoint[111]: TI201_SIG Filtrate Temperature Signal default
   		- Reset Loop : Set to 0 the DigitalPoint[112 to 149].EnableCfg
   
   -----------------------------------------------------------------------------------------------------------------------------------------------------
   	History
   		2019-DEC-24 - Merck - Q. Spindler - Initial version for Candidate Release 1.00.00.00.a
   		2020-MAR-25 - Merck - Q. Spindler - Modifications for Candidate Release 1.00.00.00.b
   					- Change the Options to enable YA17
   		2020-JUN-09 - Merck - Q. Spindler - Modifications for Candidate Release 1.00.00.00.c
   					- Remove Priority for ZSDF
   					- Change Active state to 1 for YA16
   		2020-SEP-18 - Merck - Q. Spindler - Modifications for Candidate Release 1.00.00.00.d
   					- Disable WI201_SIG alarm if ExternalWeight not used
   					- Disable TCU101_SIG alarm if ExternalTCU not used
   		2021-NOV-22 - Merck - Q. Spindler - Modifications for Candidate Release 1.01.00.00.a
   					- Add DigitalPoint[73]: YA41 Operating Time Exceeded
   		2022-SEP-22 - Actemium - J. Jaekel - Modifications for Candidate Release 1.01.00.01.a
   					- Add - DigitalPoint[111]: TI201_SIG Filtrate Temperature Signal default
   ============================================================*)
   
   (*DigitalPoint[50]: YA01 PC to PLC Com. Failure
   ============================================================*)
   DigitalPoint[50].EnableCfg := 1 ;
   DigitalPoint[50].ActiveStateCFg := 0 ;
   DigitalPoint[50].RealInputCfg := 0 ;
   DigitalPoint[50].InputAddressCfg := 50 ;
   DigitalPoint[50].AlarmCfg := 1 ;
   DigitalPoint[50].AlarmStateCfg := 1 ;
   DigitalPoint[50].OverrideCfg := 1 ;
   DigitalPoint[50].PriorityCfg := 1 ;
   DigitalPoint[50].Cond1Cfg := 1 ;
   DigitalPoint[50].Cond2Cfg := 0 ;
   DigitalPoint[50].FlashingInputCfg := 0 ;
   
   (*DigitalPoint[51]: YA02 CCP Runtime Com. Failure
   ============================================================*)
   DigitalPoint[51].EnableCfg := 1 ;
   DigitalPoint[51].ActiveStateCFg := 0 ;
   DigitalPoint[51].RealInputCfg := 0 ;
   DigitalPoint[51].InputAddressCfg := 51 ;
   DigitalPoint[51].AlarmCfg := 1 ;
   DigitalPoint[51].AlarmStateCfg := 1 ;
   DigitalPoint[51].OverrideCfg := 1 ;
   DigitalPoint[51].PriorityCfg := 1 ;
   DigitalPoint[51].Cond1Cfg := 1 ;
   DigitalPoint[51].Cond2Cfg := 0 ;
   DigitalPoint[51].FlashingInputCfg := 0 ;
   
   (*DigitalPoint[52]: YA03 Historical Data Collection Failure
   ============================================================*)
   DigitalPoint[52].EnableCfg := 1 ;
   DigitalPoint[52].ActiveStateCFg := 0 ;
   DigitalPoint[52].RealInputCfg := 0 ;
   DigitalPoint[52].InputAddressCfg := 52 ;
   DigitalPoint[52].AlarmCfg := 1 ;
   DigitalPoint[52].AlarmStateCfg := 1 ;
   DigitalPoint[52].OverrideCfg := 1 ;
   DigitalPoint[52].PriorityCfg := 1 ;
   DigitalPoint[52].Cond1Cfg := 1 ;
   DigitalPoint[52].Cond2Cfg := 0 ;
   DigitalPoint[52].FlashingInputCfg := 0 ;
   
   (*DigitalPoint[53]: YA04 Hard drive Overload
   ============================================================*)
   DigitalPoint[53].EnableCfg := 1 ;
   DigitalPoint[53].ActiveStateCFg := 1 ;
   DigitalPoint[53].RealInputCfg := 0 ;
   DigitalPoint[53].InputAddressCfg := 53 ;
   DigitalPoint[53].AlarmCfg := 1 ;
   DigitalPoint[53].AlarmStateCfg := 1 ;
   DigitalPoint[53].OverrideCfg := 1 ;
   DigitalPoint[53].PriorityCfg := 1 ;
   DigitalPoint[53].Cond1Cfg := 0 ;
   DigitalPoint[53].Cond2Cfg := 0 ;
   DigitalPoint[53].FlashingInputCfg := 0 ;
   
   (*DigitalPoint[54]: YA05 Database Overload
   ============================================================*)
   DigitalPoint[54].EnableCfg := 1 ;
   DigitalPoint[54].ActiveStateCFg := 1 ;
   DigitalPoint[54].RealInputCfg := 0 ;
   DigitalPoint[54].InputAddressCfg := 54 ;
   DigitalPoint[54].AlarmCfg := 1 ;
   DigitalPoint[54].AlarmStateCfg := 1 ;
   DigitalPoint[54].OverrideCfg := 1 ;
   DigitalPoint[54].PriorityCfg := 1 ;
   DigitalPoint[54].Cond1Cfg := 0 ;
   DigitalPoint[54].Cond2Cfg := 0 ;
   DigitalPoint[54].FlashingInputCfg := 0 ;
   
   (*DigitalPoint[55]: YA06 Node 0 Communication Failure - Smart
   ============================================================*)
   DigitalPoint[55].EnableCfg := 1 ;
   DigitalPoint[55].ActiveStateCFg := 1 ;
   DigitalPoint[55].RealInputCfg := 0;
   DigitalPoint[55].InputAddressCfg := 55 ;
   DigitalPoint[55].AlarmCfg := 1 ;
   DigitalPoint[55].AlarmStateCfg := 1 ;
   DigitalPoint[55].OverrideCfg := 1 ;
   DigitalPoint[55].PriorityCfg := 1 ;
   DigitalPoint[55].Cond1Cfg := 0 ;
   DigitalPoint[55].Cond2Cfg := 0 ;
   DigitalPoint[55].FlashingInputCfg := 0 ;
   
   (*DigitalPoint[56]: YA07 Node 0 Internal Defect - Smart
   ============================================================*)
   DigitalPoint[56].EnableCfg := 1 ;
   DigitalPoint[56].ActiveStateCFg := 1 ;
   DigitalPoint[56].RealInputCfg := 0 ;
   DigitalPoint[56].InputAddressCfg := 56 ;
   DigitalPoint[56].AlarmCfg := 1 ;
   DigitalPoint[56].AlarmStateCfg := 1 ;
   DigitalPoint[56].OverrideCfg := 1 ;
   DigitalPoint[56].PriorityCfg := 1 ;
   DigitalPoint[56].Cond1Cfg := 0 ;
   DigitalPoint[56].Cond2Cfg := 0 ;
   DigitalPoint[56].FlashingInputCfg := 0 ;
   
   (*DigitalPoint[57]: YA08 Node 1 Communication Failure - Clamshell
   ============================================================*)
   DigitalPoint[57].EnableCfg := 1 ;
   DigitalPoint[57].ActiveStateCFg := 1 ;
   DigitalPoint[57].RealInputCfg := 0 ;
   DigitalPoint[57].InputAddressCfg := 57 ;
   DigitalPoint[57].AlarmCfg := 1 ;
   DigitalPoint[57].AlarmStateCfg := 1 ;
   DigitalPoint[57].OverrideCfg := 1 ;
   DigitalPoint[57].PriorityCfg := 1 ;
   DigitalPoint[57].Cond1Cfg := 0 ;
   DigitalPoint[57].Cond2Cfg := 0 ;
   DigitalPoint[57].FlashingInputCfg := 0 ;
   
   (*DigitalPoint[58]: YA09 Node 1 Internal Defect - Clamshell
   ============================================================*)
   DigitalPoint[58].EnableCfg := 1 ;
   DigitalPoint[58].ActiveStateCFg := 1 ;
   DigitalPoint[58].RealInputCfg := 0 ;
   DigitalPoint[58].InputAddressCfg := 58 ;
   DigitalPoint[58].AlarmCfg := 1 ;
   DigitalPoint[58].AlarmStateCfg := 1 ;
   DigitalPoint[58].OverrideCfg := 1 ;
   DigitalPoint[58].PriorityCfg := 1 ;
   DigitalPoint[58].Cond1Cfg := 0 ;
   DigitalPoint[58].Cond2Cfg := 0 ;
   DigitalPoint[58].FlashingInputCfg := 0 ;
   
   (*DigitalPoint[59]: YA10 PLC Program Major Fault
   ============================================================*)
   DigitalPoint[59].EnableCfg := 1 ;
   DigitalPoint[59].ActiveStateCFg := 0 ;
   DigitalPoint[59].RealInputCfg := 0 ;
   DigitalPoint[59].InputAddressCfg := 59 ;
   DigitalPoint[59].AlarmCfg := 1 ;
   DigitalPoint[59].AlarmStateCfg := 1 ;
   DigitalPoint[59].OverrideCfg := 0 ;
   DigitalPoint[59].Priority := 1 ;
   DigitalPoint[59].PriorityCfg := 0 ;
   DigitalPoint[59].Cond1Cfg := 0 ;
   DigitalPoint[59].Cond2Cfg := 0 ;
   DigitalPoint[59].FlashingInputCfg := 0 ;
   
   (*DigitalPoint[60]: YA11 Database Corrupted
   ============================================================*)
   DigitalPoint[60].EnableCfg := 1 ;
   DigitalPoint[60].ActiveStateCFg := 1 ;
   DigitalPoint[60].RealInputCfg := 0 ;
   DigitalPoint[60].InputAddressCfg := 60 ;
   DigitalPoint[60].AlarmCfg := 1 ;
   DigitalPoint[60].AlarmStateCfg := 1 ;
   DigitalPoint[60].OverrideCfg := 1 ;
   DigitalPoint[60].PriorityCfg := 1 ;
   DigitalPoint[60].Cond1Cfg := 0 ;
   DigitalPoint[60].Cond2Cfg := 0 ;
   DigitalPoint[60].FlashingInputCfg := 0 ;
   
   (*DigitalPoint[61]: YA12 Unauthorized accesses
   ============================================================*)
   DigitalPoint[61].EnableCfg := 1 ;
   DigitalPoint[61].ActiveStateCFg := 1 ;
   DigitalPoint[61].RealInputCfg := 0 ;
   DigitalPoint[61].InputAddressCfg := 61 ;
   DigitalPoint[61].AlarmCfg := 1 ;
   DigitalPoint[61].AlarmStateCfg := 1 ;
   DigitalPoint[61].OverrideCfg := 1 ;
   DigitalPoint[61].PriorityCfg := 1 ;
   DigitalPoint[61].Cond1Cfg := 0 ;
   DigitalPoint[61].Cond2Cfg := 0 ;
   DigitalPoint[61].FlashingInputCfg := 0 ;
   
   (*DigitalPoint[62]: YA13 Tank Size Mismatch
   ============================================================*)
   IF Options.FeedTank THEN
   	DigitalPoint[62].EnableCfg := 1 ;
   	DigitalPoint[62].AlarmCfg := 1 ;
   ELSE
   	DigitalPoint[62].EnableCfg := 0 ;
   	DigitalPoint[62].AlarmCfg := 0 ;
   	DigitalPoint[62].Alarm := 0 ;
   END_IF;
   DigitalPoint[62].ActiveStateCFg := 1 ;
   DigitalPoint[62].RealInputCfg := 0 ;
   DigitalPoint[62].InputAddressCfg := 62 ;
   DigitalPoint[62].AlarmStateCfg := 1 ;
   DigitalPoint[62].OverrideCfg := 1 ;
   DigitalPoint[62].PriorityCfg := 1 ;
   DigitalPoint[62].Cond1Cfg := 0 ;
   DigitalPoint[62].Cond2Cfg := 0 ;
   DigitalPoint[62].FlashingInputCfg := 0 ;
   
   (*DigitalPoint[63]: YA14 SQL Server Write Failure
   ============================================================*)
   DigitalPoint[63].EnableCfg := 1 ;
   DigitalPoint[63].ActiveStateCFg := 0 ;
   DigitalPoint[63].RealInputCfg := 0 ;
   DigitalPoint[63].InputAddressCfg := 63 ;
   DigitalPoint[63].AlarmCfg := 1 ;
   DigitalPoint[63].AlarmStateCfg := 1 ;
   DigitalPoint[63].OverrideCfg := 0 ;
   DigitalPoint[63].PriorityCfg := 0 ;
   DigitalPoint[63].Priority := 0 ;
   DigitalPoint[63].Cond1Cfg := 0 ;
   DigitalPoint[63].Cond2Cfg := 0 ;
   DigitalPoint[63].FlashingInputCfg := 0 ;
   
   (*DigitalPoint[64]: UserNCr1 User Non Critical Alarm 1
   ============================================================*)
   DigitalPoint[64].EnableCfg := 1 ;
   DigitalPoint[64].ActiveStateCFg := 0 ;
   DigitalPoint[64].RealInputCfg := 0 ;
   DigitalPoint[64].InputAddressCfg := 64 ;
   DigitalPoint[64].AlarmCfg := 0 ;
   DigitalPoint[64].AlarmStateCfg := 0 ;
   DigitalPoint[64].OverrideCfg := 0 ;
   DigitalPoint[64].Override := 0 ;
   DigitalPoint[64].PriorityCfg := 0 ;
   DigitalPoint[64].Priority := 0 ;
   DigitalPoint[64].Cond1Cfg := 0 ;
   DigitalPoint[64].Cond2Cfg := 0 ;
   DigitalPoint[64].FlashingInputCfg := 0 ;
   
   (*DigitalPoint[65]: UserCr1 User Critical Alarm 1
   ============================================================*)
   DigitalPoint[65].EnableCfg := 1 ;
   DigitalPoint[65].ActiveStateCFg := 0 ;
   DigitalPoint[65].RealInputCfg := 0 ;
   DigitalPoint[65].InputAddressCfg := 65 ;
   DigitalPoint[65].AlarmCfg := 0 ;
   DigitalPoint[65].AlarmStateCfg := 0 ;
   DigitalPoint[65].OverrideCfg := 0 ;
   DigitalPoint[65].Override := 0 ;
   DigitalPoint[65].PriorityCfg := 0 ;
   DigitalPoint[65].Priority := 1 ;
   DigitalPoint[65].Cond1Cfg := 0 ;
   DigitalPoint[65].Cond2Cfg := 0 ;
   DigitalPoint[65].FlashingInputCfg := 0 ;
   
   (*DigitalPoint[66]: UserNCr2 User Non Critical Alarm 2
   ============================================================*)
   DigitalPoint[66].EnableCfg := 1 ;
   DigitalPoint[66].ActiveStateCFg := 0 ;
   DigitalPoint[66].RealInputCfg := 0 ;
   DigitalPoint[66].InputAddressCfg := 66 ;
   DigitalPoint[66].AlarmCfg := 0 ;
   DigitalPoint[66].AlarmStateCfg := 0 ;
   DigitalPoint[66].OverrideCfg := 0 ;
   DigitalPoint[66].Override := 0 ;
   DigitalPoint[66].PriorityCfg := 0 ;
   DigitalPoint[66].Priority := 0 ;
   DigitalPoint[66].Cond1Cfg := 0 ;
   DigitalPoint[66].Cond2Cfg := 0 ;
   DigitalPoint[66].FlashingInputCfg := 0 ;
   
   (*DigitalPoint[67]: UserCr2 User Critical Alarm 2
   ============================================================*)
   DigitalPoint[67].EnableCfg := 1 ;
   DigitalPoint[67].ActiveStateCFg := 0 ;
   DigitalPoint[67].RealInputCfg := 0 ;
   DigitalPoint[67].InputAddressCfg := 67 ;
   DigitalPoint[67].AlarmCfg := 0 ;
   DigitalPoint[67].AlarmStateCfg := 0 ;
   DigitalPoint[67].OverrideCfg := 0 ;
   DigitalPoint[67].Override := 0 ;
   DigitalPoint[67].PriorityCfg := 0 ;
   DigitalPoint[67].Priority := 1 ;
   DigitalPoint[67].Cond1Cfg := 0 ;
   DigitalPoint[67].Cond2Cfg := 0 ;
   DigitalPoint[67].FlashingInputCfg := 0 ;
   
   (*DigitalPoint[68]: ZSDF Clamshell Locking Defect
   ============================================================*)
   DigitalPoint[68].EnableCfg := 1 ;
   DigitalPoint[68].ActiveStateCFg := 1 ;
   DigitalPoint[68].RealInputCfg := 0 ;
   DigitalPoint[68].InputAddressCfg := 68 ;
   DigitalPoint[68].AlarmCfg := 1 ;
   DigitalPoint[68].AlarmStateCfg := 1 ;
   DigitalPoint[68].OverrideCfg := 1 ;
   DigitalPoint[68].PriorityCfg := 1 ;
   DigitalPoint[68].Cond1Cfg := 0 ;
   DigitalPoint[68].Cond2Cfg := 0 ;
   DigitalPoint[68].FlashingInputCfg := 0 ;
   
   (*DigitalPoint[69]: YA15 ACT350 Communication Failure
   ============================================================*)
   DigitalPoint[69].EnableCfg := 1 ;
   DigitalPoint[69].ActiveStateCFg := 1 ;
   DigitalPoint[69].RealInputCfg := 0 ;
   DigitalPoint[69].InputAddressCfg := 69 ;
   DigitalPoint[69].AlarmCfg := 1 ;
   DigitalPoint[69].AlarmStateCfg := 1 ;
   DigitalPoint[69].OverrideCfg := 1 ;
   DigitalPoint[69].PriorityCfg := 1 ;
   DigitalPoint[69].Cond1Cfg := 0 ;
   DigitalPoint[69].Cond2Cfg := 0 ;
   DigitalPoint[69].FlashingInputCfg := 0 ;
   
   (*DigitalPoint[70]: YA16 Watchdog Gateway
   ============================================================*)
   IF Options.Gateway THEN
   	DigitalPoint[70].EnableCfg := 1 ;
   	DigitalPoint[70].AlarmCfg := 1 ;
   ELSE
   	DigitalPoint[70].EnableCfg := 0 ;
   	DigitalPoint[70].AlarmCfg := 0 ;
   	DigitalPoint[70].Alarm := 0 ;
   END_IF;
   DigitalPoint[70].ActiveStateCFg := 1 ;
   DigitalPoint[70].RealInputCfg := 0 ;
   DigitalPoint[70].InputAddressCfg := 70 ;
   DigitalPoint[70].AlarmStateCfg := 0 ;
   DigitalPoint[70].OverrideCfg := 1 ;
   DigitalPoint[70].PriorityCfg := 1 ;
   DigitalPoint[70].Cond1Cfg := 0 ;
   DigitalPoint[70].Cond2Cfg := 0 ;
   DigitalPoint[70].FlashingInputCfg := 0 ;
   
   (*DigitalPoint[71]: YA17 Mobius Device Communication Failure
   ============================================================*)
   IF Options.TankPH OR Options.SingleUsePH THEN
   	DigitalPoint[71].EnableCfg := 1 ;
   	DigitalPoint[71].AlarmCfg := 1 ;
   ELSE
   	DigitalPoint[71].EnableCfg := 0 ;
   	DigitalPoint[71].AlarmCfg := 0 ;
   	DigitalPoint[71].Alarm := 0 ;
   END_IF;
   DigitalPoint[71].ActiveStateCFg := 1 ;
   DigitalPoint[71].RealInputCfg := 0 ;
   DigitalPoint[71].InputAddressCfg := 71 ;
   DigitalPoint[71].AlarmStateCfg := 1 ;
   DigitalPoint[71].OverrideCfg := 1 ;
   DigitalPoint[71].PriorityCfg := 1 ;
   DigitalPoint[71].Cond1Cfg := 0 ;
   DigitalPoint[71].Cond2Cfg := 0 ;
   DigitalPoint[71].FlashingInputCfg := 0 ;
   
   (*DigitalPoint[72]: YA18 Pump Type Mismatch
   ============================================================*)
   DigitalPoint[72].EnableCfg := 1 ;
   DigitalPoint[72].ActiveStateCFg := 1 ;
   DigitalPoint[72].RealInputCfg := 0 ;
   DigitalPoint[72].InputAddressCfg := 72 ;
   DigitalPoint[72].AlarmCfg := 1 ;
   DigitalPoint[72].AlarmStateCfg := 1 ;
   DigitalPoint[72].OverrideCfg := 1 ;
   DigitalPoint[72].PriorityCfg := 1 ;
   DigitalPoint[72].Cond1Cfg := 0 ;
   DigitalPoint[72].Cond2Cfg := 0 ;
   DigitalPoint[72].FlashingInputCfg := 0 ;
   
   (*DigitalPoint[73]: YA41 Operating Time Exceeded - Always non critical
   ============================================================*)
   DigitalPoint[73].EnableCfg := 1 ;
   DigitalPoint[73].ActiveStateCFg := 1 ;
   DigitalPoint[73].RealInputCfg := 0 ;
   DigitalPoint[73].InputAddressCfg := 73 ;
   DigitalPoint[73].AlarmCfg := 1 ;
   DigitalPoint[73].AlarmStateCfg := 1 ;
   DigitalPoint[73].OverrideCfg := 1 ;
   DigitalPoint[73].Priority := 0 ;
   DigitalPoint[73].PriorityCfg := 0 ;
   DigitalPoint[73].Cond1Cfg := 0 ;
   DigitalPoint[73].Cond2Cfg := 0 ;
   DigitalPoint[73].FlashingInputCfg := 0 ;
   
   (*Reset Loop : Set to 0 the DigitalPoint[74 to 89].EnableCfg
   ============================================================*)
   FOR Config.IndexDP := 74 to 89 by 1 do
   	DigitalPoint[Config.IndexDP].EnableCfg := 0 ;
   	DigitalPoint[Config.IndexDP].AlarmCfg := 0 ;
   	DigitalPoint[Config.IndexDP].Alarm := 0 ;
   End_for ;
   
   (*DigitalPoint[90]: AI201A_SIG Filtrate Conductivity Process Signal default
   ============================================================*)
   IF Options.FiltrateCondPH OR Options.FiltrateCondPHUV THEN
   	DigitalPoint[90].EnableCfg := 1 ;
   	DigitalPoint[90].AlarmCfg := 1 ;
   ELSE
   	DigitalPoint[90].EnableCfg := 0 ;
   	DigitalPoint[90].AlarmCfg := 0 ;
   	DigitalPoint[90].Alarm := 0 ;
   END_IF;
   DigitalPoint[90].ActiveStateCFg := 1 ;
   DigitalPoint[90].RealInputCfg := 0 ;
   DigitalPoint[90].InputAddressCfg := 90 ;
   DigitalPoint[90].AlarmStateCfg := 1 ;
   DigitalPoint[90].OverrideCfg := 1 ;
   DigitalPoint[90].PriorityCfg := 1 ;
   DigitalPoint[90].Cond1Cfg := 0 ;
   DigitalPoint[90].Cond2Cfg := 0 ;
   DigitalPoint[90].FlashingInputCfg := 0 ;
   
   (*DigitalPoint[91]: AI203_SIG Filtrate UV1 Signal default
   ============================================================*)
   IF Options.FiltrateCondPHUV THEN
   	DigitalPoint[91].EnableCfg := 1 ;
   	DigitalPoint[91].AlarmCfg := 1 ;
   ELSE
   	DigitalPoint[91].EnableCfg := 0 ;
   	DigitalPoint[91].AlarmCfg := 0 ;
   	DigitalPoint[91].Alarm := 0 ;
   END_IF;
   DigitalPoint[91].ActiveStateCFg := 1 ;
   DigitalPoint[91].RealInputCfg := 0 ;
   DigitalPoint[91].InputAddressCfg := 91 ;
   DigitalPoint[91].AlarmStateCfg := 1 ;
   DigitalPoint[91].OverrideCfg := 1 ;
   DigitalPoint[91].PriorityCfg := 1 ;
   DigitalPoint[91].Cond1Cfg := 0 ;
   DigitalPoint[91].Cond2Cfg := 0 ;
   DigitalPoint[91].FlashingInputCfg := 0 ;
   
   (*DigitalPoint[92]: AI204_SIG Filtrate UV2 Signal default
   ============================================================*)
   IF Options.FiltrateCondPHUV THEN
   	DigitalPoint[92].EnableCfg := 1 ;
   	DigitalPoint[92].AlarmCfg := 1 ;
   ELSE
   	DigitalPoint[92].EnableCfg := 0 ;
   	DigitalPoint[92].AlarmCfg := 0 ;
   	DigitalPoint[92].Alarm := 0 ;
   END_IF;
   DigitalPoint[92].ActiveStateCFg := 1 ;
   DigitalPoint[92].RealInputCfg := 0 ;
   DigitalPoint[92].InputAddressCfg := 92 ;
   DigitalPoint[92].AlarmStateCfg := 1 ;
   DigitalPoint[92].OverrideCfg := 1 ;
   DigitalPoint[92].PriorityCfg := 1 ;
   DigitalPoint[92].Cond1Cfg := 0 ;
   DigitalPoint[92].Cond2Cfg := 0 ;
   DigitalPoint[92].FlashingInputCfg := 0 ;
   
   (*DigitalPoint[93]: FI201_SIG Filtrate Flow Signal default
   ============================================================*)
   DigitalPoint[93].EnableCfg := 1 ;
   DigitalPoint[93].AlarmCfg := 1 ;
   DigitalPoint[93].ActiveStateCFg := 1 ;
   DigitalPoint[93].RealInputCfg := 0 ;
   DigitalPoint[93].InputAddressCfg := 93 ;
   DigitalPoint[93].AlarmStateCfg := 1 ;
   DigitalPoint[93].OverrideCfg := 1 ;
   DigitalPoint[93].PriorityCfg := 1 ;
   DigitalPoint[93].Cond1Cfg := 0 ;
   DigitalPoint[93].Cond2Cfg := 0 ;
   DigitalPoint[93].FlashingInputCfg := 0 ;
   
   (*DigitalPoint[94]: FI401_SIG Transfer Pump Flow Signal default
   ============================================================*)
   IF Options.TransferFlow THEN
   	DigitalPoint[94].EnableCfg := 1 ;
   	DigitalPoint[94].AlarmCfg := 1 ;
   ELSE
   	DigitalPoint[94].EnableCfg := 0 ;
   	DigitalPoint[94].AlarmCfg := 0 ;
   	DigitalPoint[94].Alarm := 0 ;
   END_IF;
   DigitalPoint[94].ActiveStateCFg := 1 ;
   DigitalPoint[94].RealInputCfg := 0 ;
   DigitalPoint[94].InputAddressCfg := 94 ;
   DigitalPoint[94].AlarmStateCfg := 1 ;
   DigitalPoint[94].OverrideCfg := 1 ;
   DigitalPoint[94].PriorityCfg := 1 ;
   DigitalPoint[94].Cond1Cfg := 0 ;
   DigitalPoint[94].Cond2Cfg := 0 ;
   DigitalPoint[94].FlashingInputCfg := 0 ;
   
   (*DigitalPoint[95]: PI601_SIG Feed Tank Pressure Signal default
   ============================================================*)
   IF Options.FeedTank THEN
   	DigitalPoint[95].EnableCfg := 1 ;
   	DigitalPoint[95].AlarmCfg := 1 ;
   ELSE
   	DigitalPoint[95].EnableCfg := 0 ;
   	DigitalPoint[95].AlarmCfg := 0 ;
   	DigitalPoint[95].Alarm := 0 ;
   END_IF;
   DigitalPoint[95].ActiveStateCFg := 1 ;
   DigitalPoint[95].RealInputCfg := 0 ;
   DigitalPoint[95].InputAddressCfg := 95 ;
   DigitalPoint[95].AlarmStateCfg := 1 ;
   DigitalPoint[95].OverrideCfg := 1 ;
   DigitalPoint[95].PriorityCfg := 1 ;
   DigitalPoint[95].Cond1Cfg := 0 ;
   DigitalPoint[95].Cond2Cfg := 0 ;
   DigitalPoint[95].FlashingInputCfg := 0 ;
   
   (*DigitalPoint[96]: WI201_SIG External Filtrate Weight Signal default
   ============================================================*)
   IF ExternalWeight THEN
   	DigitalPoint[96].AlarmCfg := 1 ;
   ELSE
   	DigitalPoint[96].AlarmCfg := 0 ;
   	DigitalPoint[96].Alarm := 0 ;
   END_IF;
   DigitalPoint[96].EnableCfg := 1 ;
   DigitalPoint[96].ActiveStateCFg := 1 ;
   DigitalPoint[96].RealInputCfg := 0 ;
   DigitalPoint[96].InputAddressCfg := 96 ;
   DigitalPoint[96].AlarmStateCfg := 1 ;
   DigitalPoint[96].OverrideCfg := 1 ;
   DigitalPoint[96].PriorityCfg := 1 ;
   DigitalPoint[96].Cond1Cfg := 0 ;
   DigitalPoint[96].Cond2Cfg := 0 ;
   DigitalPoint[96].FlashingInputCfg := 0 ;
   
   (*DigitalPoint[97]: PI001_SIG Feed Pressure Signal default
   ============================================================*)
   DigitalPoint[97].EnableCfg := 1 ;
   DigitalPoint[97].ActiveStateCFg := 1 ;
   DigitalPoint[97].RealInputCfg := 0 ;
   DigitalPoint[97].InputAddressCfg := 97 ;
   DigitalPoint[97].AlarmCfg := 1 ;
   DigitalPoint[97].AlarmStateCfg := 1 ;
   DigitalPoint[97].OverrideCfg := 1 ;
   DigitalPoint[97].PriorityCfg := 1 ;
   DigitalPoint[97].Cond1Cfg := 0 ;
   DigitalPoint[97].Cond2Cfg := 0 ;
   DigitalPoint[97].FlashingInputCfg := 0 ;
   
   (*DigitalPoint[98]: PI101_SIG Retentate Pressure Signal default
   ============================================================*)
   DigitalPoint[98].EnableCfg := 1 ;
   DigitalPoint[98].ActiveStateCFg := 1 ;
   DigitalPoint[98].RealInputCfg := 0 ;
   DigitalPoint[98].InputAddressCfg := 98 ;
   DigitalPoint[98].AlarmCfg := 1 ;
   DigitalPoint[98].AlarmStateCfg := 1 ;
   DigitalPoint[98].OverrideCfg := 1 ;
   DigitalPoint[98].PriorityCfg := 1 ;
   DigitalPoint[98].Cond1Cfg := 0 ;
   DigitalPoint[98].Cond2Cfg := 0 ;
   DigitalPoint[98].FlashingInputCfg := 0 ;
   
   (*DigitalPoint[99]: PI201_SIG Filtrate Pressure Signal default
   ============================================================*)
   DigitalPoint[99].EnableCfg := 1 ;
   DigitalPoint[99].ActiveStateCFg := 1 ;
   DigitalPoint[99].RealInputCfg := 0 ;
   DigitalPoint[99].InputAddressCfg := 99 ;
   DigitalPoint[99].AlarmCfg := 1 ;
   DigitalPoint[99].AlarmStateCfg := 1 ;
   DigitalPoint[99].OverrideCfg := 1 ;
   DigitalPoint[99].PriorityCfg := 1 ;
   DigitalPoint[99].Cond1Cfg := 0 ;
   DigitalPoint[99].Cond2Cfg := 0 ;
   DigitalPoint[99].FlashingInputCfg := 0 ;
   
   (*DigitalPoint[100]: PI401_SIG Transfer Pump Pressure Signal default
   ============================================================*)
   DigitalPoint[100].EnableCfg := 1 ;
   DigitalPoint[100].ActiveStateCFg := 1 ;
   DigitalPoint[100].RealInputCfg := 0 ;
   DigitalPoint[100].InputAddressCfg := 100 ;
   DigitalPoint[100].AlarmCfg := 1 ;
   DigitalPoint[100].AlarmStateCfg := 1 ;
   DigitalPoint[100].OverrideCfg := 1 ;
   DigitalPoint[100].PriorityCfg := 1 ;
   DigitalPoint[100].Cond1Cfg := 0 ;
   DigitalPoint[100].Cond2Cfg := 0 ;
   DigitalPoint[100].FlashingInputCfg := 0 ;
   
   (*DigitalPoint[101]: TI101_SIG Feed Tank Temperature Signal default
   ============================================================*)
   IF Options.FeedTank THEN
   	DigitalPoint[101].EnableCfg := 1 ;
   	DigitalPoint[101].AlarmCfg := 1 ;
   ELSE
   	DigitalPoint[101].EnableCfg := 0 ;
   	DigitalPoint[101].AlarmCfg := 0 ;
   	DigitalPoint[101].Alarm := 0 ;
   END_IF;
   DigitalPoint[101].ActiveStateCFg := 1 ;
   DigitalPoint[101].RealInputCfg := 0 ;
   DigitalPoint[101].InputAddressCfg := 101 ;
   DigitalPoint[101].AlarmStateCfg := 1 ;
   DigitalPoint[101].OverrideCfg := 1 ;
   DigitalPoint[101].PriorityCfg := 1 ;
   DigitalPoint[101].Cond1Cfg := 0 ;
   DigitalPoint[101].Cond2Cfg := 0 ;
   DigitalPoint[101].FlashingInputCfg := 0 ;
   
   (*DigitalPoint[102]: PCV101_SIG PCV101 Position Signal default
   ============================================================*)
   DigitalPoint[102].EnableCfg := 1 ;
   DigitalPoint[102].AlarmCfg := 1 ;
   DigitalPoint[102].ActiveStateCFg := 1 ;
   DigitalPoint[102].RealInputCfg := 0 ;
   DigitalPoint[102].InputAddressCfg := 102 ;
   DigitalPoint[102].AlarmStateCfg := 1 ;
   DigitalPoint[102].OverrideCfg := 1 ;
   DigitalPoint[102].PriorityCfg := 1 ;
   DigitalPoint[102].Cond1Cfg := 0 ;
   DigitalPoint[102].Cond2Cfg := 0 ;
   DigitalPoint[102].FlashingInputCfg := 0 ;
   
   (*DigitalPoint[103]: PCV201_SIG PCV201 Position Signal default
   ============================================================*)
   DigitalPoint[103].EnableCfg := 1 ;
   DigitalPoint[103].ActiveStateCFg := 1 ;
   DigitalPoint[103].RealInputCfg := 0 ;
   DigitalPoint[103].InputAddressCfg := 103 ;
   DigitalPoint[103].AlarmCfg := 1 ;
   DigitalPoint[103].AlarmStateCfg := 1 ;
   DigitalPoint[103].OverrideCfg := 1 ;
   DigitalPoint[103].PriorityCfg := 1 ;
   DigitalPoint[103].Cond1Cfg := 0 ;
   DigitalPoint[103].Cond2Cfg := 0 ;
   DigitalPoint[103].FlashingInputCfg := 0 ;
   
   (*DigitalPoint[104]: MIX101_SIG Mixer Speed Signal default
   ============================================================*)
   IF Options.FeedTank THEN
   	DigitalPoint[104].EnableCfg := 1 ;
   	DigitalPoint[104].AlarmCfg := 1 ;
   ELSE
   	DigitalPoint[104].EnableCfg := 0 ;
   	DigitalPoint[104].AlarmCfg := 0 ;
   	DigitalPoint[104].Alarm := 0 ;
   END_IF;
   DigitalPoint[104].ActiveStateCFg := 1 ;
   DigitalPoint[104].RealInputCfg := 0 ;
   DigitalPoint[104].InputAddressCfg := 104 ;
   DigitalPoint[104].AlarmStateCfg := 1 ;
   DigitalPoint[104].OverrideCfg := 1 ;
   DigitalPoint[104].PriorityCfg := 1 ;
   DigitalPoint[104].Cond1Cfg := 0 ;
   DigitalPoint[104].Cond2Cfg := 0 ;
   DigitalPoint[104].FlashingInputCfg := 0 ;
   
   (*DigitalPoint[105]: AI202_SIG Filtrate pH Signal default
   ============================================================*)
   IF Options.FiltrateCondPH OR Options.FiltrateCondPHUV THEN
   	DigitalPoint[105].EnableCfg := 1 ;
   	DigitalPoint[105].AlarmCfg := 1 ;
   ELSE
   	DigitalPoint[105].EnableCfg := 0 ;
   	DigitalPoint[105].AlarmCfg := 0 ;
   	DigitalPoint[105].Alarm := 0 ;
   END_IF;
   DigitalPoint[105].ActiveStateCFg := 1 ;
   DigitalPoint[105].RealInputCfg := 0 ;
   DigitalPoint[105].InputAddressCfg := 105 ;
   DigitalPoint[105].AlarmStateCfg := 1 ;
   DigitalPoint[105].OverrideCfg := 1 ;
   DigitalPoint[105].PriorityCfg := 1 ;
   DigitalPoint[105].Cond1Cfg := 0 ;
   DigitalPoint[105].Cond2Cfg := 0 ;
   DigitalPoint[105].FlashingInputCfg := 0 ;
   
   (*DigitalPoint[106]: AI101_SIG Feed Tank pH Signal default
   ============================================================*)
   IF Options.FeedTank AND Options.TankPH THEN
   	DigitalPoint[106].EnableCfg := 1 ;
   	DigitalPoint[106].AlarmCfg := 1 ;
   ELSE
   	DigitalPoint[106].EnableCfg := 0 ;
   	DigitalPoint[106].AlarmCfg := 0 ;
   	DigitalPoint[106].Alarm := 0 ;
   END_IF;
   DigitalPoint[106].ActiveStateCFg := 1 ;
   DigitalPoint[106].RealInputCfg := 0 ;
   DigitalPoint[106].InputAddressCfg := 106 ;
   DigitalPoint[106].AlarmStateCfg := 1 ;
   DigitalPoint[106].OverrideCfg := 1 ;
   DigitalPoint[106].PriorityCfg := 1 ;
   DigitalPoint[106].Cond1Cfg := 0 ;
   DigitalPoint[106].Cond2Cfg := 0 ;
   DigitalPoint[106].FlashingInputCfg := 0 ;
   
   (*DigitalPoint[107]: AI104_SIG Feed Tank Conductivity Signal default
   ============================================================*)
   IF Options.FeedTank AND Options.TankCond THEN
   	DigitalPoint[107].EnableCfg := 1 ;
   	DigitalPoint[107].AlarmCfg := 1 ;
   ELSE
   	DigitalPoint[107].EnableCfg := 0 ;
   	DigitalPoint[107].AlarmCfg := 0 ;
   	DigitalPoint[107].Alarm := 0 ;
   END_IF;
   DigitalPoint[107].ActiveStateCFg := 1 ;
   DigitalPoint[107].RealInputCfg := 0 ;
   DigitalPoint[107].InputAddressCfg := 107 ;
   DigitalPoint[107].AlarmStateCfg := 1 ;
   DigitalPoint[107].OverrideCfg := 1 ;
   DigitalPoint[107].PriorityCfg := 1 ;
   DigitalPoint[107].Cond1Cfg := 0 ;
   DigitalPoint[107].Cond2Cfg := 0 ;
   DigitalPoint[107].FlashingInputCfg := 0 ;
   
   (*DigitalPoint[108]: TCU101_SIG TCU Temperature Signal default
   ============================================================*)
   IF Options.FeedTank THEN
   	DigitalPoint[108].EnableCfg := 1 ;
   	IF ExternalTCU THEN
   		DigitalPoint[108].AlarmCfg := 1 ;
   	ELSE
   		DigitalPoint[108].AlarmCfg := 0 ;
   		DigitalPoint[108].Alarm := 0 ;
   	END_IF;
   ELSE
   	DigitalPoint[108].EnableCfg := 0 ;
   	DigitalPoint[108].AlarmCfg := 0 ;
   	DigitalPoint[108].Alarm := 0 ;
   END_IF;
   DigitalPoint[108].ActiveStateCFg := 1 ;
   DigitalPoint[108].RealInputCfg := 0 ;
   DigitalPoint[108].InputAddressCfg := 108 ;
   DigitalPoint[108].AlarmStateCfg := 1 ;
   DigitalPoint[108].OverrideCfg := 1 ;
   DigitalPoint[108].PriorityCfg := 1 ;
   DigitalPoint[108].Cond1Cfg := 0 ;
   DigitalPoint[108].Cond2Cfg := 0 ;
   DigitalPoint[108].FlashingInputCfg := 0 ;
   
   (*DigitalPoint[109]: AI201B_SIG Filtrate Conductivity Cleaning Signal default
   ============================================================*)
   IF Options.FiltrateCondPH OR Options.FiltrateCondPHUV THEN
   	DigitalPoint[109].EnableCfg := 1 ;
   	DigitalPoint[109].AlarmCfg := 1 ;
   ELSE
   	DigitalPoint[109].EnableCfg := 0 ;
   	DigitalPoint[109].AlarmCfg := 0 ;
   	DigitalPoint[109].Alarm := 0 ;
   END_IF;
   DigitalPoint[109].ActiveStateCFg := 1 ;
   DigitalPoint[109].RealInputCfg := 0 ;
   DigitalPoint[109].InputAddressCfg := 109 ;
   DigitalPoint[109].AlarmStateCfg := 1 ;
   DigitalPoint[109].OverrideCfg := 1 ;
   DigitalPoint[109].PriorityCfg := 1 ;
   DigitalPoint[109].Cond1Cfg := 0 ;
   DigitalPoint[109].Cond2Cfg := 0 ;
   DigitalPoint[109].FlashingInputCfg := 0 ;
   
   (*DigitalPoint[110]: FI101_SIG Retentate Flow Signal default
   ============================================================*)
   DigitalPoint[110].EnableCfg := 1 ;
   DigitalPoint[110].AlarmCfg := 1 ;
   DigitalPoint[110].ActiveStateCFg := 1 ;
   DigitalPoint[110].RealInputCfg := 0 ;
   DigitalPoint[110].InputAddressCfg := 110 ;
   DigitalPoint[110].AlarmStateCfg := 1 ;
   DigitalPoint[110].OverrideCfg := 1 ;
   DigitalPoint[110].PriorityCfg := 1 ;
   DigitalPoint[110].Cond1Cfg := 0 ;
   DigitalPoint[110].Cond2Cfg := 0 ;
   DigitalPoint[110].FlashingInputCfg := 0 ;
   
   (*DigitalPoint[111]: TI201_SIG Filtrate Temperature Signal default
   ============================================================*)
   IF Options.FiltrateCondPH OR Options.FiltrateCondPHUV THEN
   	DigitalPoint[111].EnableCfg := 1 ;
   	DigitalPoint[111].AlarmCfg := 1 ;
   ELSE
   	DigitalPoint[111].EnableCfg := 0 ;
   	DigitalPoint[111].AlarmCfg := 0 ;
   	DigitalPoint[111].Alarm := 0 ;
   END_IF;
   DigitalPoint[111].ActiveStateCFg := 1 ;
   DigitalPoint[111].RealInputCfg := 0 ;
   DigitalPoint[111].InputAddressCfg := 111 ;
   DigitalPoint[111].AlarmStateCfg := 1 ;
   DigitalPoint[111].OverrideCfg := 1 ;
   DigitalPoint[111].PriorityCfg := 1 ;
   DigitalPoint[111].Cond1Cfg := 0 ;
   DigitalPoint[111].Cond2Cfg := 0 ;
   DigitalPoint[111].FlashingInputCfg := 0 ;
   
   (*Reset Loop : Set to 0 the DigitalPoint[112 to 149].EnableCfg
   ============================================================*)
   FOR Config.IndexDP := 112 to 149 by 1 do
   	DigitalPoint[Config.IndexDP].EnableCfg := 0 ;
   	DigitalPoint[Config.IndexDP].AlarmCfg := 0 ;
   	DigitalPoint[Config.IndexDP].Alarm := 0 ;
   End_for ;
END_ROUTINE

ROUTINE Config_Drive   (* structured text *)
   (* ==========================================================
   	Config Drive : Configure Drive Structure (for Pumps)
   
   	List of treatments
   		- Drive[1] : Feed Pump SIC001
   		- Drive[2] : Transfer Pump SIC002
   		- Drive[3] : Mixer SIC004
   		- Reset Loop : Set to 0 the Drive[0 and 4 to 10].EnableCfg
   
   -----------------------------------------------------------------------------------------------------------------------------------------------------
   	History
   		2019-DEC-24 - Merck - Q. Spindler - Initial version for Candidate Release 1.00.00.00.a
   ============================================================*)
   
   
   (*Drive[1] : Feed Pump SIC001
   ============================================================*)
   Drive[1].EnableCfg := 1 ;
   IF Options.TFF20 THEN
   	Drive[1].OutputAddress := 8 ; // P001
   ELSE
   	Drive[1].OutputAddress := 15 ; // P003
   END_IF;
   Drive[1].InputAddress := 0 ;
   Drive[1].RunInput := 0 ;
   Drive[1].InterlockTimer.PRE := 1000 ;
   Drive[1].ReverseCfg := 0 ;
   Drive[1].DirectionAddress := 0 ;
   
   (*Drive[2] : Transfer Pump SIC002
   ============================================================*)
   Drive[2].EnableCfg := 1 ;
   Drive[2].OutputAddress := 9 ; // P002
   Drive[2].InputAddress := 0 ;
   Drive[2].RunInput := 0 ;
   Drive[2].InterlockTimer.PRE := 1000 ;
   Drive[2].ReverseCfg := 0 ;
   Drive[2].DirectionAddress := 0 ;
   
   (*Drive[3] : Mixer SIC004
   ============================================================*)
   IF Options.FeedTank THEN
   	Drive[3].EnableCfg := 1 ;
   ELSE
   	Drive[3].EnableCfg := 0 ;
   END_IF;
   Drive[3].OutputAddress := 16 ; // MIX101
   Drive[3].InputAddress := 0 ;
   Drive[3].RunInput := 0 ;
   Drive[3].InterlockTimer.PRE := 1000 ;
   Drive[3].ReverseCfg := 0 ;
   Drive[3].DirectionAddress := 0 ;
   
   (*Reset Loop : Set to 0 the Drive[0 and 4 to 10].EnableCfg
   ============================================================*)
   for Config.IndexDr := 0 to 10 by 1 do
   	if Config.IndexDr = 0 or Config.IndexDr >= 4 then
   		Drive[Config.IndexDr].EnableCfg := 0 ;
   	End_if ;
   End_for ;
END_ROUTINE

ROUTINE Config_Flowpath   (* structured text *)
   (* =======================================================================
   	Config Flowpath : Configure predifined flowpath
   
   	List of treatments
   		- Critical
   		- Common
   		- Option 1
   		- Option 2
   		- Reset Loop : Set to 0 the mask and truth of Flowpath[34 to 39]
   		- User
   		- Reset Loop : Set to 0 the mask and truth of Flowpath[45 to 60]
   		- Open All Valve (reserved)
   		- Close All Valve (reserved)
   
   -----------------------------------------------------------------------------------------------------------------------------------------------------
   	History
   		2019-DEC-24 - Merck - Q. Spindler - Initial version for Candidate Release 1.00.00.00.a
   		2020-APR-15 - Merck - Q. Spindler - Modifications for Candidate Release 1.00.00.00.b
   					- Critical Flowpath Changed (XV003 closed)
   =========================================================================*)
   
   (* Max flowpath number use as terminal value in loop
   =========================================================================*)
   FlowPathControl.MaxFlowPath := 63 ;
   
   (* Critical
   =========================================================================*)
   (* Critical *)
   
   	FlowPath[2].Mask1 := 2097151 ;
   	FlowPath[2].Mask2 := 0 ;
   	FlowPath[2].Mask3 := 0 ;
   	FlowPath[2].Mask4 := 0 ;
   	FlowPath[2].Truth1 := 387 ;
   	FlowPath[2].Truth2 := 0 ;
   	FlowPath[2].Truth3 := 0 ;
   	FlowPath[2].Truth4 := 0 ;
   
   
   (* Common
   =========================================================================*)
   
   (* Single Pass Flush (from inlet manifold) *)
   	FlowPath[3].Mask1 := 2064527 ;
   	FlowPath[3].Mask2 := 0 ;
   	FlowPath[3].Mask3 := 0 ;
   	FlowPath[3].Mask4 := 0 ;
   	FlowPath[3].Truth1 := 1114123 ;
   	FlowPath[3].Truth2 := 0 ;
   	FlowPath[3].Truth3 := 0 ;
   	FlowPath[3].Truth4 := 0 ;
   
   (* Single Pass Flush (from recycle bag) *)
   	FlowPath[4].Mask1 := 2064527 ;
   	FlowPath[4].Mask2 := 0 ;
   	FlowPath[4].Mask3 := 0 ;
   	FlowPath[4].Mask4 := 0 ;
   	FlowPath[4].Truth1 := 1114119 ;
   	FlowPath[4].Truth2 := 0 ;
   	FlowPath[4].Truth3 := 0 ;
   	FlowPath[4].Truth4 := 0 ;
   
   (* System Drain (without recycle bag) *)
   	FlowPath[5].Mask1 := 2064527 ;
   	FlowPath[5].Mask2 := 0 ;
   	FlowPath[5].Mask3 := 0 ;
   	FlowPath[5].Mask4 := 0 ;
   	FlowPath[5].Truth1 := 1900555 ;
   	FlowPath[5].Truth2 := 0 ;
   	FlowPath[5].Truth3 := 0 ;
   	FlowPath[5].Truth4 := 0 ;
   
   (* System Drain (from recycle bag) *)
   	FlowPath[6].Mask1 := 2064783 ;
   	FlowPath[6].Mask2 := 0 ;
   	FlowPath[6].Mask3 := 0 ;
   	FlowPath[6].Mask4 := 0 ;
   	FlowPath[6].Truth1 := 1900935 ;
   	FlowPath[6].Truth2 := 0 ;
   	FlowPath[6].Truth3 := 0 ;
   	FlowPath[6].Truth4 := 0 ;
   
   (* Membrane Soak *)
   	FlowPath[7].Mask1 := 2065283 ;
   	FlowPath[7].Mask2 := 0 ;
   	FlowPath[7].Mask3 := 0 ;
   	FlowPath[7].Mask4 := 0 ;
   	FlowPath[7].Truth1 := 3 ;
   	FlowPath[7].Truth2 := 0 ;
   	FlowPath[7].Truth3 := 0 ;
   	FlowPath[7].Truth4 := 0 ;
   
   (* Integrity Test *)
   	FlowPath[8].Mask1 := 2065283 ;
   	FlowPath[8].Mask2 := 0 ;
   	FlowPath[8].Mask3 := 0 ;
   	FlowPath[8].Mask4 := 0 ;
   	FlowPath[8].Truth1 := 524928 ;
   	FlowPath[8].Truth2 := 0 ;
   	FlowPath[8].Truth3 := 0 ;
   	FlowPath[8].Truth4 := 0 ;
   
   (* Recycle Bag Fill *)
   	FlowPath[9].Mask1 := 2065287 ;
   	FlowPath[9].Mask2 := 0 ;
   	FlowPath[9].Mask3 := 0 ;
   	FlowPath[9].Mask4 := 0 ;
   	FlowPath[9].Truth1 := 768 ;
   	FlowPath[9].Truth2 := 0 ;
   	FlowPath[9].Truth3 := 0 ;
   	FlowPath[9].Truth4 := 0 ;
   
   (* Recycle Bag Drain *)
   	FlowPath[10].Mask1 := 2065295 ;
   	FlowPath[10].Mask2 := 0 ;
   	FlowPath[10].Mask3 := 0 ;
   	FlowPath[10].Mask4 := 0 ;
   	FlowPath[10].Truth1 := 262149 ;
   	FlowPath[10].Truth2 := 0 ;
   	FlowPath[10].Truth3 := 0 ;
   	FlowPath[10].Truth4 := 0 ;
   
   (* Recovery Filter Flush *)
   	FlowPath[11].Mask1 := 2065295 ;
   	FlowPath[11].Mask2 := 0 ;
   	FlowPath[11].Mask3 := 0 ;
   	FlowPath[11].Mask4 := 0 ;
   	FlowPath[11].Truth1 := 131077 ;
   	FlowPath[11].Truth2 := 0 ;
   	FlowPath[11].Truth3 := 0 ;
   	FlowPath[11].Truth4 := 0 ;
   
   (* Batch UF or Membrane Recycle *)
   	FlowPath[12].Mask1 := 2065295 ;
   	FlowPath[12].Mask2 := 0 ;
   	FlowPath[12].Mask3 := 0 ;
   	FlowPath[12].Mask4 := 0 ;
   	FlowPath[12].Truth1 := 65927 ;
   	FlowPath[12].Truth2 := 0 ;
   	FlowPath[12].Truth3 := 0 ;
   	FlowPath[12].Truth4 := 0 ;
   
   (* Fed Batch UF or Diafiltration *)
   	FlowPath[13].Mask1 := 2065295 ;
   	FlowPath[13].Mask2 := 0 ;
   	FlowPath[13].Mask3 := 0 ;
   	FlowPath[13].Mask4 := 0 ;
   	FlowPath[13].Truth1 := 66439 ;
   	FlowPath[13].Truth2 := 0 ;
   	FlowPath[13].Truth3 := 0 ;
   	FlowPath[13].Truth4 := 0 ;
   
   (* Product Recovery 1&3 – Empty Recycle Bag *)
   	FlowPath[14].Mask1 := 2065295 ;
   	FlowPath[14].Mask2 := 0 ;
   	FlowPath[14].Mask3 := 0 ;
   	FlowPath[14].Mask4 := 0 ;
   	FlowPath[14].Truth1 := 131077 ;
   	FlowPath[14].Truth2 := 0 ;
   	FlowPath[14].Truth3 := 0 ;
   	FlowPath[14].Truth4 := 0 ;
   
   (* Product Recovery 2 – Empty Retentate Line *)
   	FlowPath[15].Mask1 := 2065295 ;
   	FlowPath[15].Mask2 := 0 ;
   	FlowPath[15].Mask3 := 0 ;
   	FlowPath[15].Mask4 := 0 ;
   	FlowPath[15].Truth1 := 772 ;
   	FlowPath[15].Truth2 := 0 ;
   	FlowPath[15].Truth3 := 0 ;
   	FlowPath[15].Truth4 := 0 ;
   
   (* Product Recovery 4 – Empty membranes *)
   	FlowPath[16].Mask1 := 2065283 ;
   	FlowPath[16].Mask2 := 0 ;
   	FlowPath[16].Mask3 := 0 ;
   	FlowPath[16].Mask4 := 0 ;
   	FlowPath[16].Truth1 := 131714 ;
   	FlowPath[16].Truth2 := 0 ;
   	FlowPath[16].Truth3 := 0 ;
   	FlowPath[16].Truth4 := 0 ;
   
   (* All Main Flowpath Valves Open *)
   	FlowPath[17].Mask1 := 2065283 ;
   	FlowPath[17].Mask2 := 0 ;
   	FlowPath[17].Mask3 := 0 ;
   	FlowPath[17].Mask4 := 0 ;
   	FlowPath[17].Truth1 := 2065283 ;
   	FlowPath[17].Truth2 := 0 ;
   	FlowPath[17].Truth3 := 0 ;
   	FlowPath[17].Truth4 := 0 ;
   
   (* All Main Flowpath Valves Closed *)
   	FlowPath[18].Mask1 := 2065283 ;
   	FlowPath[18].Mask2 := 0 ;
   	FlowPath[18].Mask3 := 0 ;
   	FlowPath[18].Mask4 := 0 ;
   	FlowPath[18].Truth1 := 0 ;
   	FlowPath[18].Truth2 := 0 ;
   	FlowPath[18].Truth3 := 0 ;
   	FlowPath[18].Truth4 := 0 ;
   
   (* Fill Filtrate Line (from inlet manifold) *)
   	FlowPath[19].Mask1 := 2065295 ;
   	FlowPath[19].Mask2 := 0 ;
   	FlowPath[19].Mask3 := 0 ;
   	FlowPath[19].Mask4 := 0 ;
   	FlowPath[19].Truth1 := 1081355 ;
   	FlowPath[19].Truth2 := 0 ;
   	FlowPath[19].Truth3 := 0 ;
   	FlowPath[19].Truth4 := 0 ;
   
   (* Fill Filtrate Line (from recycle bag) *)
   	FlowPath[20].Mask1 := 2065295 ;
   	FlowPath[20].Mask2 := 0 ;
   	FlowPath[20].Mask3 := 0 ;
   	FlowPath[20].Mask4 := 0 ;
   	FlowPath[20].Truth1 := 33159 ;
   	FlowPath[20].Truth2 := 0 ;
   	FlowPath[20].Truth3 := 0 ;
   	FlowPath[20].Truth4 := 0 ;
   
   (* All Source Valves Open *)
   	FlowPath[21].Mask1 := 31868 ;
   	FlowPath[21].Mask2 := 0 ;
   	FlowPath[21].Mask3 := 0 ;
   	FlowPath[21].Mask4 := 0 ;
   	FlowPath[21].Truth1 := 31864 ;
   	FlowPath[21].Truth2 := 0 ;
   	FlowPath[21].Truth3 := 0 ;
   	FlowPath[21].Truth4 := 0 ;
   
   (* All Source Valves Closed *)
   	FlowPath[22].Mask1 := 31864 ;
   	FlowPath[22].Mask2 := 0 ;
   	FlowPath[22].Mask3 := 0 ;
   	FlowPath[22].Mask4 := 0 ;
   	FlowPath[22].Truth1 := 0 ;
   	FlowPath[22].Truth2 := 0 ;
   	FlowPath[22].Truth3 := 0 ;
   	FlowPath[22].Truth4 := 0 ;
   
   (* Option 1
   =========================================================================*)
   
   (* Feed Source Open *)
   	FlowPath[23].Mask1 := 31744 ;
   	FlowPath[23].Mask2 := 0 ;
   	FlowPath[23].Mask3 := 0 ;
   	FlowPath[23].Mask4 := 0 ;
   	FlowPath[23].Truth1 := 1024 ;
   	FlowPath[23].Truth2 := 0 ;
   	FlowPath[23].Truth3 := 0 ;
   	FlowPath[23].Truth4 := 0 ;
   
   (* Buffer Source Open *)
   	FlowPath[24].Mask1 := 31744 ;
   	FlowPath[24].Mask2 := 0 ;
   	FlowPath[24].Mask3 := 0 ;
   	FlowPath[24].Mask4 := 0 ;
   	FlowPath[24].Truth1 := 2048 ;
   	FlowPath[24].Truth2 := 0 ;
   	FlowPath[24].Truth3 := 0 ;
   	FlowPath[24].Truth4 := 0 ;
   
   (* Caustic Source Open *)
   	FlowPath[25].Mask1 := 31744 ;
   	FlowPath[25].Mask2 := 0 ;
   	FlowPath[25].Mask3 := 0 ;
   	FlowPath[25].Mask4 := 0 ;
   	FlowPath[25].Truth1 := 4096 ;
   	FlowPath[25].Truth2 := 0 ;
   	FlowPath[25].Truth3 := 0 ;
   	FlowPath[25].Truth4 := 0 ;
   
   (* Water Source Open *)
   	FlowPath[26].Mask1 := 31744 ;
   	FlowPath[26].Mask2 := 0 ;
   	FlowPath[26].Mask3 := 0 ;
   	FlowPath[26].Mask4 := 0 ;
   	FlowPath[26].Truth1 := 8192 ;
   	FlowPath[26].Truth2 := 0 ;
   	FlowPath[26].Truth3 := 0 ;
   	FlowPath[26].Truth4 := 0 ;
   
   (* Air Source Open *)
   	FlowPath[27].Mask1 := 31744 ;
   	FlowPath[27].Mask2 := 0 ;
   	FlowPath[27].Mask3 := 0 ;
   	FlowPath[27].Mask4 := 0 ;
   	FlowPath[27].Truth1 := 16384 ;
   	FlowPath[27].Truth2 := 0 ;
   	FlowPath[27].Truth3 := 0 ;
   	FlowPath[27].Truth4 := 0 ;
   
   (* Option 2
   =========================================================================*)
   
   (* Feed Source Open - Xfer line *)
   	FlowPath[28].Mask1 := 7168 ;
   	FlowPath[28].Mask2 := 0 ;
   	FlowPath[28].Mask3 := 0 ;
   	FlowPath[28].Mask4 := 0 ;
   	FlowPath[28].Truth1 := 1024 ;
   	FlowPath[28].Truth2 := 0 ;
   	FlowPath[28].Truth3 := 0 ;
   	FlowPath[28].Truth4 := 0 ;
   
   (* Buffer Source Open - Xfer line *)
   	FlowPath[29].Mask1 := 7168 ;
   	FlowPath[29].Mask2 := 0 ;
   	FlowPath[29].Mask3 := 0 ;
   	FlowPath[29].Mask4 := 0 ;
   	FlowPath[29].Truth1 := 2048 ;
   	FlowPath[29].Truth2 := 0 ;
   	FlowPath[29].Truth3 := 0 ;
   	FlowPath[29].Truth4 := 0 ;
   
   (* Air Source Open - Xfer line *)
   	FlowPath[30].Mask1 := 7168 ;
   	FlowPath[30].Mask2 := 0 ;
   	FlowPath[30].Mask3 := 0 ;
   	FlowPath[30].Mask4 := 0 ;
   	FlowPath[30].Truth1 := 4096 ;
   	FlowPath[30].Truth2 := 0 ;
   	FlowPath[30].Truth3 := 0 ;
   	FlowPath[30].Truth4 := 0 ;
   (*
   
   (* Caustic Source Open - Feed line *)
   	FlowPath[31].Mask1 := 124 ;
   	FlowPath[31].Mask2 := 0 ;
   	FlowPath[31].Mask3 := 0 ;
   	FlowPath[31].Mask4 := 0 ;
   	FlowPath[31].Truth1 := 24 ;
   	FlowPath[31].Truth2 := 0 ;
   	FlowPath[31].Truth3 := 0 ;
   	FlowPath[31].Truth4 := 0 ;
   (*
   
   (* Water Source Open - Feed line *)
   	FlowPath[32].Mask1 := 124 ;
   	FlowPath[32].Mask2 := 0 ;
   	FlowPath[32].Mask3 := 0 ;
   	FlowPath[32].Mask4 := 0 ;
   	FlowPath[32].Truth1 := 40 ;
   	FlowPath[32].Truth2 := 0 ;
   	FlowPath[32].Truth3 := 0 ;
   	FlowPath[32].Truth4 := 0 ;
   (*
   
   (* Buffer/Air Source Open - Feed line *)
   	FlowPath[33].Mask1 := 124 ;
   	FlowPath[33].Mask2 := 0 ;
   	FlowPath[33].Mask3 := 0 ;
   	FlowPath[33].Mask4 := 0 ;
   	FlowPath[33].Truth1 := 72 ;
   	FlowPath[33].Truth2 := 0 ;
   	FlowPath[33].Truth3 := 0 ;
   	FlowPath[33].Truth4 := 0 ;
   
   (*Reset Loop : Set to 0 the Flowpath[34 to 39]
   ============================================================*)
   FOR Config.IndexFlowpath := 34 to 39 by 1 do
   	FlowPath[Config.IndexFlowpath].Mask1 := 0 ;
   	FlowPath[Config.IndexFlowpath].Mask2 := 0 ;
   	FlowPath[Config.IndexFlowpath].Mask3 := 0 ;
   	FlowPath[Config.IndexFlowpath].Mask4 := 0 ;
   	FlowPath[Config.IndexFlowpath].Truth1 := 0 ;
   	FlowPath[Config.IndexFlowpath].Truth2 := 0 ;
   	FlowPath[Config.IndexFlowpath].Truth3 := 0 ;
   	FlowPath[Config.IndexFlowpath].Truth4 := 0 ;
   	FlowPath[Config.IndexFlowpath].Status := 0 ;
   End_for ;
   
   
   (* User
   =========================================================================*)
   (* Flowpath from 30 to 34 are reserved for User *)
   
   
   (*Reset Loop : Set to 0 the Flowpath[45 to 60]
   ============================================================*)
   FOR Config.IndexFlowpath := 45 to 60 by 1 do
   	FlowPath[Config.IndexFlowpath].Mask1 := 0 ;
   	FlowPath[Config.IndexFlowpath].Mask2 := 0 ;
   	FlowPath[Config.IndexFlowpath].Mask3 := 0 ;
   	FlowPath[Config.IndexFlowpath].Mask4 := 0 ;
   	FlowPath[Config.IndexFlowpath].Truth1 := 0 ;
   	FlowPath[Config.IndexFlowpath].Truth2 := 0 ;
   	FlowPath[Config.IndexFlowpath].Truth3 := 0 ;
   	FlowPath[Config.IndexFlowpath].Truth4 := 0 ;
   	FlowPath[Config.IndexFlowpath].Status := 0 ;
   End_for ;
   
   
   (* Open All Valve (reserved)
   =========================================================================*)
   (* Open All Valve *)
   FlowPath[61].Mask1 := -1 ;
   FlowPath[61].Mask2 := 0 ;
   FlowPath[61].Mask3 := 0 ;
   FlowPath[61].Mask4 := 0 ;
   FlowPath[61].Truth1 := -1 ;
   FlowPath[61].Truth2 := 0 ;
   FlowPath[61].Truth3 := 0 ;
   FlowPath[61].Truth4 := 0 ;
   
   (* Close All Valve (reserved)
   =========================================================================*)
   (* Close All Valve *)
   FlowPath[62].Mask1 := -1 ;
   FlowPath[62].Mask2 := 0 ;
   FlowPath[62].Mask3 := 0 ;
   FlowPath[62].Mask4 := 0 ;
   FlowPath[62].Truth1 := 0 ;
   FlowPath[62].Truth2 := 0 ;
   FlowPath[62].Truth3 := 0 ;
   FlowPath[62].Truth4 := 0 ;
   
END_ROUTINE
